(* IEC 61131-3 sources: daoli-st-library/DL_MathData (part 8) *)

(* ---- FC_DL_AngleLerpShort.st ---- *)
(*==============================================================================
 * 名称 : FC_DL_AngleLerpShort —— 两角度最短弧线性插值（跨 0/360 正确）
 * 分类 / 前缀 / 版本 : DL_MathData / FC_DL_ / 1.0.0
 * 溯源 : 开源语义参考（OSCAT/AixOCAT 族，MIT）或 clean-room IEC 实现，未复制源码
 * 平台 : 纯 IEC 61131-3
 * 功能说明 : 沿 fA→fB 最短弧做线性插值：先求 fB-fA 的最短弧差 d∈[-180,180)，
 *            结果 = fA + fT*d，再归一到 [0,360)。fT=0 得 fA 方向，fT=1 得 fB
 *            方向；跨 0/360（如 350°→10°）走 +20° 短弧而非 -340° 长弧。
 *            边界处理：fT 越界 [0,1] 钳位使用（不置故障，属容错钳位）；任一
 *            输入非有限（NaN/±Inf）置 eErr 返回 0.0；|fA|>1.0E12 置 eErr。
 * 错误码 : 16#0001_1B02 = 输入非有限（NaN/±Inf）或角度量超安全量程 ±1.0E12
 *          eErr=0 且 bValid=TRUE 表示返回值可用
 * 状态机 : R6 标注 N/A（纯函数无顺序状态，以本节替代 ELSE 兜底）
 * 红线 : R1/R2/R3 ✓ 零全局/零IO/纯IEC ｜ R4 ✓ 非有限拦截/钳位/量程防护 ｜ R10 ✓ 标准转换 ｜ R11 ✓ 分号收尾 ｜ R15 ✓ 无保留字撞名
 * 修订记录 : 2026-11-23 v1.0.0 首次入库（R76）
 *============================================================================*)
FUNCTION FC_DL_AngleLerpShort : LREAL
VAR_INPUT
    fA : LREAL;    // 插值起点角 [度] / interpolation start angle in degrees
    fB : LREAL;    // 插值终点角 [度] / interpolation end angle in degrees
    fT : LREAL;    // 插值比例 0..1，越界钳位 [无量纲] / interpolation ratio, clamped into [0,1]
END_VAR
VAR_OUTPUT
    eErr   : UDINT;    // 故障码，0=正常，1B02=输入非有限或超量程 / error code
    bError : BOOL;     // TRUE=本件发生故障 / TRUE when fault occurred
    bValid : BOOL;     // TRUE=返回值可用 / TRUE when return value is usable
END_VAR
VAR
    _d : LREAL;        // fA→fB 最短弧差 [度] / shortest-arc diff from A to B
    _n : LREAL;        // 整圈数（TRUNC 截断）[圈] / whole turns via truncation
    _t : LREAL;        // 钳位后的插值比例 [无量纲] / clamped ratio
    _r : LREAL;        // 插值中间结果 [度] / interpolated raw result
END_VAR

FC_DL_AngleLerpShort := 0.0;                 // 返回值预设 0.0 / preset return to zero
eErr   := 16#0000_0000;                      // 故障码清零 / clear error code
bError := FALSE;                             // 故障标志清零 / clear error flag
bValid := TRUE;                              // 预设输出可用 / preset valid flag

IF (fA <> fA) OR ((fA - fA) <> (fA - fA))    // fA 非有限 / fA is NaN or infinite
   OR (fB <> fB) OR ((fB - fB) <> (fB - fB)) // fB 非有限 / fB is NaN or infinite
   OR (fT <> fT) OR ((fT - fT) <> (fT - fT)) // fT 非有限 / fT is NaN or infinite
   OR (ABS(fA) > 1.0E12) OR (ABS(fB) > 1.0E12) THEN    // 角度量超安全量程 / beyond safe range
    eErr   := 16#0001_1B02;                  // 置故障码 / set error code
    bError := TRUE;                          // 置故障标志 / set error flag
    bValid := FALSE;                         // 返回值不可用 / return not usable
    RETURN;                                  // 返回 0.0 / return zero
END_IF

_t := fT;                                    // 取比例 / take ratio
IF _t < 0.0 THEN _t := 0.0; END_IF           // 下界钳位 / clamp lower bound
IF _t > 1.0 THEN _t := 1.0; END_IF           // 上界钳位 / clamp upper bound

_d := fB - fA;                               // 原始差值 / raw difference
_d := _d - 360.0 * TRUNC(_d / 360.0);        // 整圈截断缩圈 / strip whole turns
IF _d >= 180.0 THEN                          // 上越界修正 / fix upper overflow
    _d := _d - 360.0;                        // 减一整圈 / subtract one turn
END_IF
IF _d < -180.0 THEN                          // 下越界修正 / fix lower overflow
    _d := _d + 360.0;                        // 加一整圈 / add one turn
END_IF

_r := fA + _t * _d;                          // 沿最短弧插值 / interpolate along shortest arc
_r := _r - 360.0 * TRUNC(_r / 360.0);        // 归一缩圈 / normalize by stripping turns
IF _r < 0.0 THEN                             // 负角修正 / fix negative angle
    _r := _r + 360.0;                        // 加一整圈 / add one turn
END_IF

FC_DL_AngleLerpShort := _r;                  // 回写 [0,360) 插值结果 / write back result

END_FUNCTION

(* ---- FC_DL_AngleQuadrant.st ---- *)
(*==============================================================================
 * 名称 : FC_DL_AngleQuadrant —— 角度象限判定（0..3）与坐标轴命中标志
 * 分类 / 前缀 / 版本 : DL_MathData / FC_DL_ / 1.0.0
 * 溯源 : 开源语义参考（OSCAT/AixOCAT 族，MIT）或 clean-room IEC 实现，未复制源码
 * 平台 : 纯 IEC 61131-3
 * 功能说明 : 将输入角归一到 [0,360) 后判定象限：0=[0,90) 1=[90,180)
 *            2=[180,270) 3=[270,360)。归一角恰为 0/90/180/270（容差
 *            1.0E-9，浮点禁用 = 直接比较）时 bOnAxis=TRUE，象限取该轴线
 *            后一侧区间编号（0°→0、90°→1、180°→2、270°→3）。
 *            边界处理：输入非有限（NaN/±Inf）或 |角|>1.0E12 置 eErr 返回 0。
 * 错误码 : 16#0001_1B03 = 输入非有限（NaN/±Inf）或角度量超安全量程 ±1.0E12
 *          eErr=0 且 bValid=TRUE 表示象限与轴标志均可用
 * 状态机 : R6 标注 N/A（纯函数无顺序状态，以本节替代 ELSE 兜底）
 * 红线 : R1/R2/R3 ✓ 零全局/零IO/纯IEC ｜ R4 ✓ 非有限拦截/浮点容差比较 ｜ R10 ✓ 标准转换 ｜ R11 ✓ 分号收尾 ｜ R15 ✓ 无保留字撞名
 * 修订记录 : 2026-11-23 v1.0.0 首次入库（R76）
 *============================================================================*)
FUNCTION FC_DL_AngleQuadrant : INT
VAR_INPUT
    fAngle : LREAL;    // 输入角（任意实数，内部归一）[度] / input angle, normalized internally
END_VAR
VAR_OUTPUT
    bOnAxis : BOOL;    // TRUE=归一角命中 0/90/180/270（容差 1.0E-9）/ TRUE when on axis within 1.0E-9
    eErr    : UDINT;   // 故障码，0=正常，1B03=输入非有限或超量程 / error code
    bError  : BOOL;    // TRUE=本件发生故障 / TRUE when fault occurred
    bValid  : BOOL;    // TRUE=象限与轴标志可用 / TRUE when outputs are usable
END_VAR
VAR
    _r : LREAL;        // 归一后的角 [度] / normalized angle
    _n : LREAL;        // 整圈数（TRUNC 截断）[圈] / whole turns via truncation
END_VAR

FC_DL_AngleQuadrant := 0;                    // 象限预设 0 / preset quadrant to zero
bOnAxis := FALSE;                            // 轴标志预设 FALSE / preset on-axis to FALSE
eErr    := 16#0000_0000;                     // 故障码清零 / clear error code
bError  := FALSE;                            // 故障标志清零 / clear error flag
bValid  := TRUE;                             // 预设输出可用 / preset valid flag

IF (fAngle <> fAngle) OR ((fAngle - fAngle) <> (fAngle - fAngle))    // 非有限 / NaN or infinite
   OR (ABS(fAngle) > 1.0E12) THEN            // 超安全量程 / beyond safe range
    eErr   := 16#0001_1B03;                  // 置故障码 / set error code
    bError := TRUE;                          // 置故障标志 / set error flag
    bValid := FALSE;                         // 输出不可用 / outputs not usable
    RETURN;                                  // 返回 0 / return zero
END_IF

_r := fAngle;                                // 取输入角 / take input
_r := _r - 360.0 * TRUNC(_r / 360.0);        // 整圈截断缩圈 / strip whole turns
IF _r < 0.0 THEN                             // 负角修正 / fix negative angle
    _r := _r + 360.0;                        // 加一整圈，得 [0,360) / add one turn
END_IF

IF ABS(_r - 0.0) < 1.0E-9                    // 轴线 0°（含容差）/ on axis 0 deg
   OR ABS(_r - 90.0) < 1.0E-9                // 轴线 90°（含容差）/ on axis 90 deg
   OR ABS(_r - 180.0) < 1.0E-9               // 轴线 180°（含容差）/ on axis 180 deg
   OR ABS(_r - 270.0) < 1.0E-9 THEN          // 轴线 270°（含容差）/ on axis 270 deg
    bOnAxis := TRUE;                         // 置轴线命中标志 / set on-axis flag
END_IF

IF _r >= 270.0 THEN                          // [270,360) 第 4 象限 / quadrant 4
    FC_DL_AngleQuadrant := 3;                // 象限码 3 / quadrant code 3
ELSIF _r >= 180.0 THEN                       // [180,270) 第 3 象限 / quadrant 3
    FC_DL_AngleQuadrant := 2;                // 象限码 2 / quadrant code 2
ELSIF _r >= 90.0 THEN                        // [90,180) 第 2 象限 / quadrant 2
    FC_DL_AngleQuadrant := 1;                // 象限码 1 / quadrant code 1
ELSE                                         // [0,90) 第 1 象限 / quadrant 1
    FC_DL_AngleQuadrant := 0;                // 象限码 0 / quadrant code 0
END_IF

END_FUNCTION

(* ---- FC_DL_AngleReflect.st ---- *)
(*==============================================================================
 * 名称 : FC_DL_AngleReflect —— 关于轴线角 fAxis 的镜像反射（结果 [0,360)）
 * 分类 / 前缀 / 版本 : DL_MathData / FC_DL_ / 1.0.0
 * 溯源 : 开源语义参考（OSCAT/AixOCAT 族，MIT）或 clean-room IEC 实现，未复制源码
 * 平台 : 纯 IEC 61131-3
 * 功能说明 : 求入射角 fAngle 关于镜像轴 fAxis 的反射角：r = 2*fAxis - fAngle
 *            （数值语义恒正确，含跨 0°/360° 情形），归一到 [0,360)。
 *            例：轴 45°、入射 10° → 反射 80°；轴 0°、入射 350° → 反射 10°。
 *            边界处理：任一输入非有限（NaN/±Inf）或 |量|>1.0E12 置 eErr 返回 0.0。
 * 错误码 : 16#0001_1B07 = 输入非有限（NaN/±Inf）或角度量超安全量程 ±1.0E12
 *          eErr=0 且 bValid=TRUE 表示返回值可用
 * 状态机 : R6 标注 N/A（纯函数无顺序状态，以本节替代 ELSE 兜底）
 * 红线 : R1/R2/R3 ✓ 零全局/零IO/纯IEC ｜ R4 ✓ 非有限拦截/量程防护 ｜ R10 ✓ 标准转换 ｜ R11 ✓ 分号收尾 ｜ R15 ✓ 无保留字撞名
 * 修订记录 : 2026-11-23 v1.0.0 首次入库（R76）
 *============================================================================*)
FUNCTION FC_DL_AngleReflect : LREAL
VAR_INPUT
    fAngle : LREAL;    // 入射角 [度] / incident angle in degrees
    fAxis  : LREAL;    // 镜像轴角 [度] / mirror axis angle in degrees
END_VAR
VAR_OUTPUT
    eErr   : UDINT;    // 故障码，0=正常，1B07=输入非有限或超量程 / error code
    bError : BOOL;     // TRUE=本件发生故障 / TRUE when fault occurred
    bValid : BOOL;     // TRUE=返回值可用 / TRUE when return value is usable
END_VAR
VAR
    _r : LREAL;        // 反射角中间值 [度] / reflected raw angle
END_VAR

FC_DL_AngleReflect := 0.0;                   // 返回值预设 0.0 / preset return to zero
eErr   := 16#0000_0000;                      // 故障码清零 / clear error code
bError := FALSE;                             // 故障标志清零 / clear error flag
bValid := TRUE;                              // 预设输出可用 / preset valid flag

IF (fAngle <> fAngle) OR ((fAngle - fAngle) <> (fAngle - fAngle))    // fAngle 非有限 / NaN or infinite
   OR (fAxis <> fAxis) OR ((fAxis - fAxis) <> (fAxis - fAxis))        // fAxis 非有限 / NaN or infinite
   OR (ABS(fAngle) > 1.0E12) OR (ABS(fAxis) > 1.0E12) THEN            // 角度量超安全量程 / beyond safe range
    eErr   := 16#0001_1B07;                  // 置故障码 / set error code
    bError := TRUE;                          // 置故障标志 / set error flag
    bValid := FALSE;                         // 返回值不可用 / return not usable
    RETURN;                                  // 返回 0.0 / return zero
END_IF

_r := 2.0 * fAxis - fAngle;                  // 关于轴镜像反射 / reflect about axis
_r := _r - 360.0 * TRUNC(_r / 360.0);        // 整圈截断缩圈 / strip whole turns
IF _r < 0.0 THEN                             // 负角修正 / fix negative angle
    _r := _r + 360.0;                        // 加一整圈，得 [0,360) / add one turn
END_IF

FC_DL_AngleReflect := _r;                    // 回写 [0,360) 反射角 / write back reflection

END_FUNCTION

(* ---- FC_DL_AngleToCompass.st ---- *)
(*==============================================================================
 * 名称 : FC_DL_AngleToCompass —— 方位角转 16 方位码（0=北，顺时针）与 8 方位码
 * 分类 / 前缀 / 版本 : DL_MathData / FC_DL_ / 1.0.0
 * 溯源 : 开源语义参考（OSCAT/AixOCAT 族，MIT）或 clean-room IEC 实现，未复制源码
 * 平台 : 纯 IEC 61131-3
 * 功能说明 : 将方位角归一到 [0,360) 后按每扇区 22.5° 映射到 16 方位码
 *            0..15（0=北、4=东、8=南、12=西，顺时针），并以 45° 扇区同步
 *            给出 8 方位码 nBand 0..7（0=北、2=东、4=南、6=西），供下游
 *            粗分级直接使用。扇区中心对齐：加半扇区 11.25°/22.5° 后取整。
 *            边界处理：输入非有限（NaN/±Inf）或 |角|>1.0E12 置 eErr 返回 0。
 * 错误码 : 16#0001_1B05 = 输入非有限（NaN/±Inf）或角度量超安全量程 ±1.0E12
 *          eErr=0 且 bValid=TRUE 表示两码均可用
 * 状态机 : R6 标注 N/A（纯函数无顺序状态，以本节替代 ELSE 兜底）
 * 红线 : R1/R2/R3 ✓ 零全局/零IO/纯IEC ｜ R4 ✓ 非有限拦截/量程防护 ｜ R10 ✓ 标准转换 ｜ R11 ✓ 分号收尾 ｜ R15 ✓ 无保留字撞名
 * 修订记录 : 2026-11-23 v1.0.0 首次入库（R76）
 *============================================================================*)
FUNCTION FC_DL_AngleToCompass : INT
VAR_INPUT
    fAngle : LREAL;    // 方位角（0=北，顺时针为正）[度] / bearing angle, clockwise from north
END_VAR
VAR_OUTPUT
    nBand  : INT;      // 8 方位码 0..7（0=北）/ 8-point compass code
    eErr   : UDINT;    // 故障码，0=正常，1B05=输入非有限或超量程 / error code
    bError : BOOL;     // TRUE=本件发生故障 / TRUE when fault occurred
    bValid : BOOL;     // TRUE=两码均可用 / TRUE when both codes are usable
END_VAR
VAR
    _r    : LREAL;     // 归一后的方位角 [度] / normalized bearing
    _n16  : LREAL;     // 16 扇区整数值 / 16-sector integer value
    _n8   : LREAL;     // 8 扇区整数值 / 8-sector integer value
END_VAR

FC_DL_AngleToCompass := 0;                   // 16 码预设 0（北）/ preset 16-code to north
nBand := 0;                                  // 8 码预设 0（北）/ preset 8-code to north
eErr  := 16#0000_0000;                       // 故障码清零 / clear error code
bError:= FALSE;                              // 故障标志清零 / clear error flag
bValid:= TRUE;                               // 预设输出可用 / preset valid flag

IF (fAngle <> fAngle) OR ((fAngle - fAngle) <> (fAngle - fAngle))    // 非有限 / NaN or infinite
   OR (ABS(fAngle) > 1.0E12) THEN            // 超安全量程 / beyond safe range
    eErr   := 16#0001_1B05;                  // 置故障码 / set error code
    bError := TRUE;                          // 置故障标志 / set error flag
    bValid := FALSE;                         // 输出不可用 / outputs not usable
    RETURN;                                  // 返回 0 / return north codes
END_IF

_r := fAngle;                                // 取输入角 / take input
_r := _r - 360.0 * TRUNC(_r / 360.0);        // 整圈截断缩圈 / strip whole turns
IF _r < 0.0 THEN                             // 负角修正 / fix negative angle
    _r := _r + 360.0;                        // 加一整圈，得 [0,360) / add one turn
END_IF

_n16 := TRUNC((_r + 11.25) / 22.5);          // 16 扇区中心对齐取整 / 16-sector center-aligned
_n8  := TRUNC((_r + 22.5) / 45.0);           // 8 扇区中心对齐取整 / 8-sector center-aligned

FC_DL_AngleToCompass := DINT_TO_INT(LREAL_TO_DINT(_n16) MOD 16);    // 折回 0..15 / fold into 0..15
nBand := DINT_TO_INT(LREAL_TO_DINT(_n8) MOD 8);           // 折回 0..7 / fold into 0..7

END_FUNCTION

(* ---- FC_DL_AngleTolInside.st ---- *)
(*==============================================================================
 * 名称 : FC_DL_AngleTolInside —— 角度容差窗判定（fCenter ± fTol，跨 0° 正确）
 * 分类 / 前缀 / 版本 : DL_MathData / FC_DL_ / 1.0.0
 * 溯源 : 开源语义参考（OSCAT/AixOCAT 族，MIT）或 clean-room IEC 实现，未复制源码
 * 平台 : 纯 IEC 61131-3
 * 功能说明 : 判定 fAngle 是否落在 fCenter ± fTol 的圆周窗内：取 fAngle-fCenter
 *            的最短弧差 d∈[-180,180)（天然跨 0°/360° 正确），当 |d| <= fTol
 *            判在内。窗宽 >180° 时窗覆盖超过半圆，仍按最短弧口径判定。
 *            边界处理：fTol<0 判参数非法（置 eErr 返回 FALSE）；任一角度输入
 *            非有限（NaN/±Inf）或 |角|>1.0E12 置 eErr 返回 FALSE。
 * 错误码 : 16#0001_1B06 = fTol 为负（容差非法），或角度输入非有限 / 超安全量程 ±1.0E12
 *          eErr=0 且 bValid=TRUE 表示判定结论可用
 * 状态机 : R6 标注 N/A（纯函数无顺序状态，以本节替代 ELSE 兜底）
 * 红线 : R1/R2/R3 ✓ 零全局/零IO/纯IEC ｜ R4 ✓ 非有限拦截/浮点容差比较 ｜ R10 ✓ 标准转换 ｜ R11 ✓ 分号收尾 ｜ R15 ✓ 无保留字撞名
 * 修订记录 : 2026-11-23 v1.0.0 首次入库（R76）
 *============================================================================*)
FUNCTION FC_DL_AngleTolInside : BOOL
VAR_INPUT
    fAngle  : LREAL;   // 被判定角 [度] / angle under test in degrees
    fCenter : LREAL;   // 窗中心角 [度] / window center angle in degrees
    fTol    : LREAL;   // 容差半窗宽，须 >=0 [度] / tolerance half-width, must be >= 0
END_VAR
VAR_OUTPUT
    eErr   : UDINT;    // 故障码，0=正常，1B06=参数非法或非有限 / error code
    bError : BOOL;     // TRUE=本件发生故障 / TRUE when fault occurred
    bValid : BOOL;     // TRUE=判定结论可用 / TRUE when verdict is usable
END_VAR
VAR
    _d : LREAL;        // 最短弧差 [度] / shortest-arc diff
END_VAR

FC_DL_AngleTolInside := FALSE;               // 判定预设 FALSE / preset verdict to FALSE
eErr   := 16#0000_0000;                      // 故障码清零 / clear error code
bError := FALSE;                             // 故障标志清零 / clear error flag
bValid := TRUE;                              // 预设输出可用 / preset valid flag

IF fTol < 0.0 THEN                           // 容差为负：参数非法 / negative tolerance invalid
    eErr   := 16#0001_1B06;                  // 置参数非法码 / set invalid-parameter code
    bError := TRUE;                          // 置故障标志 / set error flag
    bValid := FALSE;                         // 结论不可用 / verdict not usable
    RETURN;                                  // 返回 FALSE / return FALSE
END_IF

IF (fAngle <> fAngle) OR ((fAngle - fAngle) <> (fAngle - fAngle))     // fAngle 非有限 / NaN or infinite
   OR (fCenter <> fCenter) OR ((fCenter - fCenter) <> (fCenter - fCenter))   // fCenter 非有限 / NaN or infinite
   OR (fTol <> fTol) OR ((fTol - fTol) <> (fTol - fTol))               // fTol 非有限 / NaN or infinite
   OR (ABS(fAngle) > 1.0E12) OR (ABS(fCenter) > 1.0E12) THEN           // 角度量超安全量程 / beyond safe range
    eErr   := 16#0001_1B06;                  // 置故障码 / set error code
    bError := TRUE;                          // 置故障标志 / set error flag
    bValid := FALSE;                         // 结论不可用 / verdict not usable
    RETURN;                                  // 返回 FALSE / return FALSE
END_IF

_d := fAngle - fCenter;                      // 原始差值 / raw difference
_d := _d - 360.0 * TRUNC(_d / 360.0);        // 整圈截断缩圈 / strip whole turns
IF _d >= 180.0 THEN                          // 上越界修正 / fix upper overflow
    _d := _d - 360.0;                        // 减一整圈 / subtract one turn
END_IF
IF _d < -180.0 THEN                          // 下越界修正 / fix lower overflow
    _d := _d + 360.0;                        // 加一整圈 / add one turn
END_IF

IF ABS(_d) <= fTol THEN                      // 最短弧差落在容差窗内 / diff inside tolerance window
    FC_DL_AngleTolInside := TRUE;            // 判在内 / verdict inside
END_IF

END_FUNCTION

(* ---- FC_DL_AngleUnwrapStep.st ---- *)
(*==============================================================================
 * 名称 : FC_DL_AngleUnwrapStep —— 增量解卷绕（跨多圈连续跟踪，步进 [-180,180)）
 * 分类 / 前缀 / 版本 : DL_MathData / FC_DL_ / 1.0.0
 * 溯源 : 开源语义参考（OSCAT/AixOCAT 族，MIT）或 clean-room IEC 实现，未复制源码
 * 平台 : 纯 IEC 61131-3
 * 功能说明 : 编码器增量解卷绕：取 fRaw-fPrev 的最短弧差作为本拍步进
 *            fStep∈[-180,180)，返回 fAccum + fStep 的累计角（不卷绕、跨多圈
 *            连续跟踪）。调用方须把返回值与 fStep 存为下一拍的 fAccum/fPrev。
 *            边界处理：任一输入非有限（NaN/±Inf）或 |量|>1.0E12 置 eErr
 *            返回 fAccum 原值（冻结本拍步进，不引入伪增量）。
 * 错误码 : 16#0001_1B08 = 输入非有限（NaN/±Inf）或角度量超安全量程 ±1.0E12
 *          eErr=0 且 bValid=TRUE 表示步进与累计角均可用
 * 状态机 : R6 标注 N/A（纯函数无顺序状态，跨拍状态由调用方持有，以本节替代 ELSE 兜底）
 * 红线 : R1/R2/R3 ✓ 零全局/零IO/纯IEC ｜ R4 ✓ 非有限拦截/量程防护 ｜ R10 ✓ 标准转换 ｜ R11 ✓ 分号收尾 ｜ R15 ✓ 无保留字撞名
 * 修订记录 : 2026-11-23 v1.0.0 首次入库（R76）
 *============================================================================*)
FUNCTION FC_DL_AngleUnwrapStep : LREAL
VAR_INPUT
    fRaw   : LREAL;    // 本拍原始角 [度] / raw angle of this cycle
    fPrev  : LREAL;    // 上一拍原始角（调用方持有）[度] / previous raw angle, caller-held
    fAccum : LREAL;    // 累计角（调用方持有）[度] / accumulated angle, caller-held
END_VAR
VAR_OUTPUT
    fStep  : LREAL;    // 本拍步进 [-180,180) [度] / step of this cycle within [-180,180)
    eErr   : UDINT;    // 故障码，0=正常，1B08=输入非有限或超量程 / error code
    bError : BOOL;     // TRUE=本件发生故障 / TRUE when fault occurred
    bValid : BOOL;     // TRUE=步进与累计角可用 / TRUE when step and result are usable
END_VAR
VAR
    _d : LREAL;        // 本拍原始差值 [度] / raw delta of this cycle
END_VAR

fStep := 0.0;                                // 步进预设 0.0 / preset step to zero
eErr   := 16#0000_0000;                      // 故障码清零 / clear error code
bError := FALSE;                             // 故障标志清零 / clear error flag
bValid := TRUE;                              // 预设输出可用 / preset valid flag
FC_DL_AngleUnwrapStep := fAccum;             // 返回值预设为累计角原值 / preset return to accum

IF (fRaw <> fRaw) OR ((fRaw - fRaw) <> (fRaw - fRaw))      // fRaw 非有限 / NaN or infinite
   OR (fPrev <> fPrev) OR ((fPrev - fPrev) <> (fPrev - fPrev))   // fPrev 非有限 / NaN or infinite
   OR (fAccum <> fAccum) OR ((fAccum - fAccum) <> (fAccum - fAccum))  // fAccum 非有限 / NaN or infinite
   OR (ABS(fRaw) > 1.0E12) OR (ABS(fPrev) > 1.0E12) THEN     // 角度量超安全量程 / beyond safe range
    eErr   := 16#0001_1B08;                  // 置故障码 / set error code
    bError := TRUE;                          // 置故障标志 / set error flag
    bValid := FALSE;                         // 输出不可用 / outputs not usable
    RETURN;                                  // 冻结本拍，返回 fAccum 原值 / freeze, return accum unchanged
END_IF

_d := fRaw - fPrev;                          // 本拍原始差值 / raw delta
_d := _d - 360.0 * TRUNC(_d / 360.0);        // 整圈截断缩圈 / strip whole turns
IF _d >= 180.0 THEN                          // 上越界修正（取短弧步进）/ fix upper overflow
    _d := _d - 360.0;                        // 减一整圈 / subtract one turn
END_IF
IF _d < -180.0 THEN                          // 下越界修正 / fix lower overflow
    _d := _d + 360.0;                        // 加一整圈 / add one turn
END_IF

fStep := _d;                                 // 回写本拍步进 / write back step
FC_DL_AngleUnwrapStep := fAccum + _d;        // 累计角连续跟踪（不卷绕）/ accumulate unwrapped

END_FUNCTION

(* ---- FC_DL_AnodizeFilmThicknessCalc.st ---- *)
(*
  Component : FC_DL_AnodizeFilmThicknessCalc
  Category  : DL_MathData
  Type      : FC
  Complexity: C1
  VERSION   : v1.0.0
  功能      : 阳极氧化膜厚-电量换算：按法拉第定律由电量密度与膜密度算膜厚 μm，并按电流密度反算达目标膜厚所需时间。
  开源溯源  : 道莅原创 clean-room 自研（无外部代码引用）｜License: MIT
  边界条件  : ① 膜密度、摩尔质量、转移电子数须 > 1e-9，效率须在 (0,100] % 内，否则返回哨兵 -1；
              ② 反算时间需电流密度 > 1e-9，电流密度为 0 时时间回 0（不下发 inf）；
              ③ 量纲链：g/dm² ÷ g/cm³ = cm³/dm²，除 dm² 面积 100 cm² 得 cm 厚，再乘 1e4 得 μm。
*)
FUNCTION FC_DL_AnodizeFilmThicknessCalc : REAL
VAR_INPUT
    fChgDensAsDm2 : REAL;   (* 电量密度 [A·s/dm²] Charge density *)
    fMolarMassGmol: REAL;   (* 氧化物摩尔质量 [g/mol] Oxide molar mass *)
    fDensityGcm3  : REAL;   (* 膜层密度 [g/cm³] Film density *)
    nElectrons    : INT;    (* 反应转移电子数 [个] Transferred electrons *)
    fEffPct       : REAL;   (* 电流效率 [%] Current efficiency *)
    fCurrDensADm2 : REAL;   (* 电流密度 [A/dm²] Current density *)
    fThickTargetUm: REAL;   (* 目标膜厚 [μm] Target film thickness *)
END_VAR
VAR_OUTPUT
    fFilmUm        : REAL;  (* 膜厚 [μm] Film thickness *)
    fMassGdm2      : REAL;  (* 单位面积氧化膜质量 [g/dm²] Film mass per area *)
    fTimeForTargetS: REAL;  (* 达目标膜厚所需时间 [s] Time to reach target thickness *)
    xValid         : BOOL;  (* 计算有效性标志 [-] Calculation valid flag *)
END_VAR
VAR CONSTANT
    DL_EPS      : REAL := 1.0E-9;   (* 除零判定容差 [无量纲] Divide-by-zero tolerance *)
    DL_FARADAY  : REAL := 96485.332;(* 法拉第常数 [C/mol] Faraday constant *)
    DL_CM_PER_DM: REAL := 100.0;    (* dm² 对应 cm² 数 [cm²/dm²] cm2 per dm2 *)
    DL_PCT_BASE : REAL := 100.0;    (* 百分比基准 [%] Percent base *)
    DL_UM_PER_CM: REAL := 10000.0;  (* 厘米转微米系数 [μm/cm] Micrometres per centimetre *)
    DL_ZERO     : REAL := 0.0;      (* 零常量 [无量纲] Zero constant *)
END_VAR
VAR
    fEffUnit : REAL;   (* 效率折算系数 [-] Efficiency as fraction *)
    fMoles   : REAL;   (* 单位面积反应摩尔数 [mol/dm²] Moles per area *)
END_VAR
(* 出口预置：四出口统一预置 *)
fFilmUm := 0.0; fMassGdm2 := 0.0; fTimeForTargetS := 0.0; xValid := FALSE;
(* 非有限拦截：自反判 NaN，自身差值判 Inf *)
IF (fChgDensAsDm2 <> fChgDensAsDm2) OR ((fChgDensAsDm2 - fChgDensAsDm2) <> 0.0)
   OR (fMolarMassGmol <> fMolarMassGmol) OR ((fMolarMassGmol - fMolarMassGmol) <> 0.0)
   OR (fDensityGcm3 <> fDensityGcm3) OR ((fDensityGcm3 - fDensityGcm3) <> 0.0)
   OR (fEffPct <> fEffPct) OR ((fEffPct - fEffPct) <> 0.0)
   OR (fCurrDensADm2 <> fCurrDensADm2) OR ((fCurrDensADm2 - fCurrDensADm2) <> 0.0) THEN
    FC_DL_AnodizeFilmThicknessCalc := -1.0;  (* 哨兵 -1：输入非有限 / Sentinel -1 non-finite *)
    RETURN;
END_IF
(* 组态域闸：膜密度、摩尔质量、转移电子数、效率、电量密度非负 *)
IF (fDensityGcm3 <= DL_EPS) OR (fMolarMassGmol <= DL_EPS) OR (nElectrons < 1)
   OR (fEffPct <= DL_ZERO) OR (fEffPct > DL_PCT_BASE) OR (fChgDensAsDm2 < DL_ZERO) THEN
    FC_DL_AnodizeFilmThicknessCalc := -1.0;  (* 哨兵 -1：组态非法 / Sentinel -1 bad config *)
    RETURN;
END_IF
fEffUnit := fEffPct / DL_PCT_BASE;             (* 效率折算 [-] / Efficiency as fraction *)
(* 单位面积摩尔数：n = q / (z·F)，电量密度为 C/dm² *)
fMoles := fChgDensAsDm2 / (INT_TO_REAL(nElectrons) * DL_FARADAY);
(* 单位面积质量：m = n·M [g/dm²]，乘效率得实际成膜量 *)
fMassGdm2 := fMoles * fMolarMassGmol * fEffUnit;
(* 厚度换算：g/dm² ÷ g/cm³ = cm³/dm²，除 100 cm² 得 cm，再乘 1e4 得 μm *)
fFilmUm := (fMassGdm2 / fDensityGcm3) / DL_CM_PER_DM * DL_UM_PER_CM;
(* 反算时间：t = 目标膜厚 / (电流密度 × 单位电量膜厚系数)，电流密度为 0 时回 0 *)
IF (fCurrDensADm2 > DL_EPS) AND (fThickTargetUm > DL_ZERO) THEN
    fTimeForTargetS := fThickTargetUm * INT_TO_REAL(nElectrons) * DL_FARADAY * fDensityGcm3
                       / (fCurrDensADm2 * fMolarMassGmol * fEffUnit * DL_CM_PER_DM);
END_IF
xValid := TRUE;                                (* 链路有效 / Chain valid *)
FC_DL_AnodizeFilmThicknessCalc := fFilmUm;     (* 返回膜厚 [μm] / Return film thickness *)
END_FUNCTION

(* ---- FC_DL_ArrayCumSumLreal.st ---- *)
(*
    FC_DL_ArrayCumSumLreal —— LREAL 数组前缀累计序列 + 总和出口（统计线）
    ------------------------------------------------------------------
    组件名称  : FC_DL_ArrayCumSumLreal
    分类      : DL_MathData / Statistics
    前缀      : FC_DL_
    版本      : 1.0.0
    溯源      : 借鉴组织 —— T2-1 LGF · Math（统计线，矩阵行 157）：仅借鉴
                「前缀累计 / 累计序列输出」公开功能定义；clean-room 声明 ——
                零代码行复制，判据链 / 码位 / 钳位与拒绝口径 100% 自有；
                累加内核为 IEC 61131-3 标准算术的道莅防御性实现。
    平台      : 纯 IEC 61131-3（WHILE + LREAL 算术），无内建函数依赖，
                CODESYS 3.5 / TwinCAT 3 / InoProShop / Machine Expert 通用
    作者      : 道莅代码库 · PLC编程专家（R72 构建轮 · 批 1 · 序号 3）
    ------------------------------------------------------------------
    功能说明  : 对有效样本数 nCount 个 LREAL 输入计算前缀累计序列
                afOut[i] = Σ afIn[1..i]（i = 1..nCount），并给总和出口
                fTotal = afOut[nCount]。真实工况：能耗 / 产量累计曲线、
                按片批次余量推演、OEE 累计谱。量纲随输入（m³ / kWh / 件 等），
                本件不解释量纲。
                判据链顺序：
                ① nCount 域闸：0 → 信息级空出口（fTotal = 0，afOut 不触碰，
                   bValid = TRUE）；> 数组上界 → 钳位照算 + 信息级；
                ② 逐元素非有限闸（两遍扫描第一遍，R151 闸全枚举）：**遇非有限
                   样本整体拒绝**（保守口径：部分累计会污染下游余量判断，
                   出故障级码，afOut 零写入）；
                ③ 循环累加（WHILE 带 DL_CUM_GUARD 防死锁计数器，两遍各自独立
                   计数）+ 写前下标双检；
                ④ 溢出面：累计 > 1E30 → 置 bTruncated 中断累加（保留至上一
                   有效前缀），信息级声明口径；非有限中间量同判（差值自反 +
                   自反双判，R79）。
                浮点判等禁用 =（红线 5）：本件无浮点相等比较。
    错误码    : 16#0002_3902 nCount = 0，空出口（fTotal = 0，bValid = TRUE）
                            —— 信息级，不置 bError（R45）
                16#0002_3903 nCount > 数组上界，已钳位照算 —— 信息级，值可用
                16#0002_3904 样本非有限或循环守卫越限（整体拒绝，afOut 零写入，
                            返回 FALSE）—— 故障级
                16#0002_3905 累计超 1E30 上界，已置 bTruncated 中断累加（保留
                            至上一有效前缀，bValid = TRUE）—— 信息级
                加码反证句（R90）：3902/3903/3905 均有独立输出观测面
                （3902 由 nCount=0 请求 + 空出口唯一对应；3903 由钳位行为 +
                部分结果唯一对应；3905 由 bTruncated 专位唯一对应），互不可
                由现有输出组合还原，故各立一码。
    码位总账  : 16#0002_3902 用 ｜ 16#0002_3903 用 ｜ 16#0002_3904 用 ｜
                16#0002_3905 用
    状态机    : N/A —— 纯函数无状态，无 CASE 可写，非法状态不可能出现
    边界与披露: 一 无定时器 / 无沿检测实例，周期安全规则 N/A；WHILE 双循环
                   各配 DL_CUM_GUARD 守卫（160 > 上界 128，正常不触发），
                   守卫越限并入 3904 故障级（结构性不可达防御收口）；
                二 零全局变量、零 VAR_EXTERNAL、零物理地址；
                三 域闸逐项点名（R272）：afIn[1..nEff] 全部元素纳入非有限闸；
                   nCount 域闸覆盖 0 / 上界两端点（各推一条向量）；
                四 数组写前下标双检（红线 2）：(nI >= 1) AND (nI <= DL_CUM_NMAX)
                   显式兜底；下标 > nCount 的 afOut 元素不被本件触碰；
                五 除法面：无（零除法，零除零面）；
                六 与 FC_DL_ArraySumLreal（DL_MathData）分工互引：后者只出
                   总和（可零拷贝、非有限剔除口径），本件输出**完整前缀序列**
                   （须写入调用方数组、整体拒绝口径），非变体，分工写死。
    验收向量  : V1 afIn = [1,2,3]，nCount = 3 → afOut = [1,3,6]，fTotal = 6；
                V2 nCount = 0 → 空出口 3902，fTotal = 0，afOut 不触碰；
                V3 nCount = 200（> 128）→ 钳位照算 3903；
                V4 afIn[2] = NaN → 3904 故障级，afOut 零写入；
                V5 累计越 1E30 → bTruncated = TRUE + 3905。
                算法已证（脚本）：未跑 ｜ 编译器已证（三平台）：未跑
    修订记录  : 2026-11-23 v1.0.0 首次入库（R72 构建轮 · 批 1 · 序号 3）
*)
FUNCTION FC_DL_ArrayCumSumLreal : BOOL
VAR_INPUT
    nCount    : UDINT;                     (* 有效样本数，[个]，0 = 空出口，超上界钳位照算 / the valid sample count *)
END_VAR
VAR_IN_OUT
    afIn      : ARRAY[1..DL_CUM_NMAX] OF LREAL;  (* 输入样本数组，[量纲随输入]，下标 1 起 / the input samples, unit follows the caller *)
    afOut     : ARRAY[1..DL_CUM_NMAX] OF LREAL;  (* 前缀累计序列出口，[量纲随输入]，afOut[i] = Σ afIn[1..i] / the prefix cumulative output *)
END_VAR
VAR_OUTPUT
    fTotal     : LREAL;                    (* 总和出口 = afOut[nCount]（截断时为最后有效前缀），[量纲随输入] / the total outlet *)
    bTruncated : BOOL;                     (* 累计越 1E30 上界截断标志 / the truncation flag *)
    bValid     : BOOL;                     (* 输出可用标志，故障级为 FALSE / the outputs usable flag *)
    bError     : BOOL;                     (* 故障标志，仅故障级码置位（R45 配对）/ the fault flag *)
    nInfoCode  : UDINT;                    (* 信息 / 错误码，0 = 正常 / the info or error id *)
END_VAR
VAR CONSTANT
    DL_CUM_NMAX  : INT  := 128;            (* 数组上界（两数组维度必须与本常量一致）[个] / the array upper bound, both arrays must match *)
    DL_CUM_NMAXU : UDINT := 128;           (* 数组上界的 UDINT 影子（nCount 域闸同口径比较用）[个] / the UDINT shadow of the bound *)
    DL_CUM_CAP   : LREAL := 1.0E30;        (* 累计幅值上界（截断口径）[量纲随输入] / the cumulative magnitude cap *)
    DL_CUM_GUARD : INT  := 160;            (* 循环守卫上限（> 上界 128，正常不触发）[次] / the loop guard limit *)
    DL_CUM_ZERO  : LREAL := 0.0;           (* 零哨兵 [量纲随输入] / the zero sentinel *)
    DL_CUM_ONE   : INT  := 1;              (* 游标步进与下界常量 [个] / the cursor step and lower bound *)
END_VAR
VAR
    nEff    : INT;                         (* 钳位后的有效样本数 [个] / the effective clamped count *)
    nI      : INT;                         (* 数组游标 [个] / the array cursor *)
    nGuard  : INT;                         (* 循环守卫计数器 [次] / the loop guard counter *)
    fRun    : LREAL;                       (* 累加器 [量纲随输入] / the running accumulator *)
    bFinOk  : BOOL;                        (* 第一遍有限性扫描结论 / the pass one finiteness verdict *)
    bStop   : BOOL;                        (* 第二遍截断中止标志 / the pass two truncation stop flag *)
    bSmpFin : BOOL;                        (* 当前样本有限性中间结论 / the per sample finiteness temporary *)
END_VAR

// 段 1｜返回值与状态预置（统一出口预置，R256）/ segment 1, preset the return and the status
FC_DL_ArrayCumSumLreal := FALSE;         // 故障缺省返回不可用 / the fault default is unusable
fTotal     := DL_CUM_ZERO;               // 总和出口预置零 / preset the total to zero
bTruncated := FALSE;                     // 截断标志预清零 / preset the truncation flag false
bValid     := FALSE;                     // 可用标志预清零 / preset the usable flag false
bError     := FALSE;                     // 故障标志预清零 / preset the fault flag false
nInfoCode  := 0;                         // 码位预置无错 / preset the code to zero
nEff    := 0;                            // 有效数预置零 / preset the effective count zero
nI      := 0;                            // 游标预置零 / preset the cursor zero
nGuard  := 0;                            // 守卫预置零 / preset the guard zero
fRun    := DL_CUM_ZERO;                  // 累加器清零 / clear the accumulator
bFinOk  := TRUE;                         // 有限性结论预置通过 / preset the finiteness verdict pass
bStop   := FALSE;                        // 截断标志预清零 / preset the stop flag false
bSmpFin := TRUE;                         // 样本有限性预置通过 / preset the per sample verdict pass

// 段 2｜nCount 域闸（0 = 空出口，超界 = 钳位照算，两端点向量）/ segment 2, the count domain gate
IF nCount = 0 THEN                       // 空请求：信息级空出口（afOut 不触碰）/ an empty request, the empty outlet
    nInfoCode := 16#0002_3902;           // 信息级：空出口 / info level: the empty outlet
    bError := FALSE;                     // 信息级不置故障（R45）/ info level never raises a fault
    bValid := TRUE;                      // 空出口按契约可用 / the empty outlet usable by contract
    FC_DL_ArrayCumSumLreal := TRUE;      // 照算完成（空）/ the pass complete, empty
    RETURN;                              // 结构早退 / structural exit
END_IF
IF nCount > DL_CUM_NMAXU THEN            // 请求超数组上界：钳位照算 / the request over the bound, clamped
    nInfoCode := 16#0002_3903;           // 信息级：已钳位照算 / info level: clamped
    nEff := DL_CUM_NMAX;                 // 钳到上界 / clamp to the bound
ELSE                                     // 域内请求 / the in domain request
    nEff := UDINT_TO_DINT(nCount);       // 降位转换（已证 <= 128，无回绕面）/ the narrowing conversion proven safe
END_IF

// 段 3｜第一遍：逐元素非有限扫描（整体拒绝口径，闸前零写入）/ segment 3, the pass one finiteness scan
nI     := DL_CUM_ONE;                    // 游标从下标 1 起 / the cursor from index one
nGuard := 0;                            // 守卫清零 / clear the guard
WHILE (nI <= nEff) AND (nGuard < DL_CUM_GUARD) DO // 守卫内扫描 / the scan inside the guard
    IF (nI >= DL_CUM_ONE) AND (nI <= DL_CUM_NMAX) THEN // 写前读前下标双检（红线 2）/ the index double check
        bSmpFin := NOT ((afIn[nI] <> afIn[nI]) OR ((afIn[nI] - afIn[nI]) <> 0.0)); // 自反 + 差值自反双判（R79）/ the reflexive pair test
        IF NOT bSmpFin THEN              // 非有限样本命中 / a non finite sample hit
            bFinOk := FALSE;             // 整体拒绝结论 / the overall reject verdict
            nI := nEff + DL_CUM_ONE;     // 跳出扫描（守卫内合法退出）/ break the scan legally
        END_IF
    END_IF
    nI := nI + DL_CUM_ONE;               // 游标推进 / advance the cursor
    nGuard := nGuard + DL_CUM_ONE;       // 守卫推进 / advance the guard
END_WHILE
IF (NOT bFinOk) OR (nGuard >= DL_CUM_GUARD) THEN // 非有限命中或守卫越限 / a hit or a guard overflow
    nInfoCode := 16#0002_3904;           // 故障级：样本序列不可信整体拒绝（守卫越限为结构性不可达防御收口）/ fault level: the samples untrusted
    bError := TRUE;                      // R45 配对置故障标志 / paired with the fault flag
    bValid := FALSE;                     // 输出不可用 / the outputs unusable
    FC_DL_ArrayCumSumLreal := FALSE;     // 拒绝返回 / the reject return
    RETURN;                              // 结构早退（afOut 保持零写入）/ exit with afOut untouched
END_IF

// 段 4｜第二遍：前缀累计与写出口（截断口径：累计 > 1E30 中断累加）/ segment 4, the pass two prefix accumulation
nI     := DL_CUM_ONE;                    // 游标复位 / reset the cursor
nGuard := 0;                             // 守卫复位 / reset the guard
WHILE (nI <= nEff) AND (nGuard < DL_CUM_GUARD) AND (NOT bStop) DO // 守卫与截断双出口 / the loop with both exits
    IF (nI >= DL_CUM_ONE) AND (nI <= DL_CUM_NMAX) THEN // 写前下标双检（红线 2）/ the index double check
        fRun := fRun + afIn[nI];         // 前缀累加（样本已过第一遍闸）/ the prefix accumulation
        IF (fRun <> fRun) OR ((fRun - fRun) <> 0.0) OR (fRun > DL_CUM_CAP) THEN // 溢出面：非有限中间量或越上界 / the overflow surface
            bTruncated := TRUE;          // 置截断标志 / raise the truncation flag
            nInfoCode := 16#0002_3905;   // 信息级：已截断（优先级高于钳位码 3903，声明口径）/ info level: truncated, overriding the clamp code
            bStop := TRUE;               // 中断累加（保留至上一有效前缀）/ stop the accumulation
        ELSE                             // 前缀有效 / the prefix valid
            afOut[nI] := fRun;           // 写前缀出口 / write the prefix outlet
        END_IF
    END_IF
    nI := nI + DL_CUM_ONE;               // 游标推进 / advance the cursor
    nGuard := nGuard + DL_CUM_ONE;       // 守卫推进 / advance the guard
END_WHILE

// 段 5｜正常出口 / segment 5, the normal outlet
fTotal := fRun;                          // 总和出口 = 最后有效前缀 / the total outlet, the last valid prefix
bError := FALSE;                         // 信息级不置故障（双保险）/ info level never raises a fault, second line
bValid := TRUE;                          // 输出可用 / the outputs usable
FC_DL_ArrayCumSumLreal := TRUE;          // 照算完成 / the pass complete
END_FUNCTION

(* ---- FC_DL_ArrayDiffSummary.st ---- *)
(*==============================================================================
 * 组件名称 (Component)  : FC_DL_ArrayDiffSummary
 * 所属子库 (Sublibrary) : DL_MathData
 * 归属目录 (Directory)  : C:\Library\DL_MathData
 * 当前版本 (Version)    : 1.0.1
 * 组件分类 (Category)   : 函数（FUNCTION）· 纯函数 · 双数组逐项容差比对
 * 兼容性   (Platform)   : CODESYS 3.5 / TwinCAT 3 / 汇川 InoProShop / 施耐德
 *                         Machine Expert；仅用 Standard.library 的 ABS，无实例依赖
 * 功能一句话 (Summary)  : 两组实数数组按统一绝对容差逐项比对，输出超差项数、首个
 *                         超差下标、最大绝对偏差及其下标与一致性结论。
 * 功能描述 (Function)   : 配方回读、双通道冗余比对、视觉参数下发校验三类场景，
 *                         现场只判「有差异」却定位不到第几项、差多少；用等号判等
 *                         又会因浮点误差把合格品报成不合格。本件一次扫描给出
 *                         计数、首个位置、最大偏差位置三个定位量，维修工直接翻表。
 * 与既有件边界 (Boundary): FC_DL_SearchMinMax 在单数组内找极值；FC_DL_ArraySearchFirst
 *                         在单数组内按判据找首个命中；本件是双数组逐项配对比较，
 *                         输出统计族，三者职责互斥，不存在覆盖关系。
 * 设计要点 (Key notes)  : ① 容差先取绝对值再钳到最小容差，杜绝「容差为零把纯浮点
 *                           噪声全判超差」的静默失效；
 *                         ② 非数与非有限值前置拦截：该项直接计为超差且不参与最大
 *                           偏差竞争，防止无穷大污染统计结果；
 *                         ③ 最大偏差并列时取先出现者，保证结果可复现；
 *                         ④ 单趟循环完成全部判定，无嵌套循环、无排序、无中间数组；
 *                         ⑤ 纯函数：无内部状态，同入参同结果，可重入。
 * 开源溯源 (Origin)     : 来源标签 lgf-comparator。LGF 为免费闭源发布的公开函数库
 *                         手册，本件仅借鉴其比较器组把「数组批量比较」与「容差窗口」
 *                         分成两个子域的分类骨架；许可证按其发布方条款仅作分类参考，
 *                         本件零代码行、零注释引用，属 clean-room 独立实现。统计口径
 *                         （最大偏差及其下标）为本库自有，LGF 批量比较不输出该量。
 * 码位说明 (Codes)      : 本件独占信息级码段 16#0001_0134 到 16#0001_0135，纯函数
 *                         无锁存面故不占故障级码；与 MathData 既有 0101 到 0124
 *                         及同轮 0125 到 013C 求差为空。
 *                         0134 项数越界已钳位 ｜ 0135 容差非法已回退。
 * 依赖说明 (Depends)    : 无 DL_ 内部依赖；仅 Standard.library 的 ABS。
 * 契约前置条件 (Contract): 函数内无法探测数组实际长度，「nCount 不得大于调用方实际
 *                         数组长度」由调用方负责，组态时须与装载行数绑定。
 * 红线自检 (Redline)    : 零全局变量表依赖 ｜ 零外部变量声明 ｜ 零物理地址
 *                         纯 IEC 61131-3 ｜ 浮点无等号判等，全部走容差 ｜ 无除法
 *                         数组下标先钳位后使用 ｜ 循环带守卫 ｜ 全变量双语同行注释
 * 修订历史 (Revision)   : 2026-11-15  v1.0.0  首版入库（Round 12 · 双数组比对族）
 *                         2026-11-15  v1.0.1  终审定点修复 A-D04：两项有限值相减仍可能
 *                         溢出为无穷（同号异号近满量程），原实现会让该偏差直接参与最大
 *                         偏差竞争并把 fMaxDev 污染成无穷；补「偏差本身超有限上限即按非
 *                         有限处置、不参与竞争」判据，兑现设计要点②的承诺
 *============================================================================*)

(*==============================================================================
 * 比对示意 (Comparison picture)：
 *   期望 10.0 / 20.0 / 30.0，实际 10.0 / 20.005 / 30.2，容差 0.01
 *   第 2 项偏差 0.005 在容差内，合格，但仍是目前最大偏差
 *   第 3 项偏差 0.2 超出容差，超差计数加一，并顶替最大偏差
 *   最终：超差一项、首个超差下标 3、最大偏差 0.2 落在下标 3、不相等
 *   若把实际第 2 项置为非数，该项计为超差且不参与最大偏差竞争
 *============================================================================*)

FUNCTION FC_DL_ArrayDiffSummary : BOOL
VAR_IN_OUT
    afExpected : ARRAY[1..64] OF REAL;   // 期望值数组，基准侧，只读不写 [工程单位] / Expected reference array, read only
    afActual   : ARRAY[1..64] OF REAL;   // 实际值数组，回读侧，只读不写 [工程单位] / Actual readback array, read only
END_VAR
VAR_INPUT
    nCount  : INT := 1;                  // 参与比对项数 [项]，域 1 到 64，越界钳位 / Item count, 1 to 64, clamped
    fAbsTol : REAL := 0.01;              // 统一绝对容差 [工程单位]，负值取绝对值 / Absolute tolerance, negative values folded to positive
END_VAR
VAR_OUTPUT
    nDiffCount   : INT;                  // 超差项数 [项] / Number of out of tolerance items
    nFirstDiffIdx : INT;                 // 首个超差项下标，0 表示无超差 [索引] / First out of tolerance index, zero when none
    fMaxDev      : REAL;                 // 最大绝对偏差值，只统计有限项 [工程单位] / Maximum absolute deviation over finite items
    nMaxDevIdx   : INT;                  // 最大偏差所在下标，0 表示未计算 [索引] / Index of the maximum deviation
    bEqual       : BOOL;                 // 全部项在容差内且无非有限值为真 / All items within tolerance and finite
    bNonFinite   : BOOL;                 // 出现过非数或非有限项为真 / NaN or infinity encountered
    uErrorId     : UDINT;                // 事件码，0 表示无事件 / Event code, zero means none
    bValid       : BOOL;                 // 项数与容差落在可服务域内为真，容差回退不否定结果 / Count and tolerance serviceable, a tolerance fallback does not void the result
END_VAR
VAR
    nCountUse : INT;                     // 生效项数，钳位后的值 [项] / Effective item count after clamping
    fTolUse   : REAL;                    // 生效容差，已取绝对值并钳到最小容差 [工程单位] / Effective tolerance after normalisation
    fDev      : REAL;                    // 单项绝对偏差 [工程单位] / Per item absolute deviation
    fA        : REAL;                    // 当前期望值快照 [工程单位] / Expected value snapshot
    fB        : REAL;                    // 当前实际值快照 [工程单位] / Actual value snapshot
    bFinA     : BOOL;                    // 期望值有限性判定结果 / Expected value finiteness
    bFinB     : BOOL;                    // 实际值有限性判定结果 / Actual value finiteness
    nGuard    : DINT;                    // 循环守卫计数，防遍历失控 [次] / Loop guard counter
    i         : INT;                     // 遍历索引，1 起 [索引] / Loop index, one based
END_VAR
VAR CONSTANT
    DL_ITEM_MAX   : INT := 64;          // 项数上限 [项] / Item count limit
    DL_GUARD_MAX  : DINT := 128;        // 循环守卫上限，两倍于项数上限故正常不触发 [次] / Loop guard limit, twice the item limit
    DL_I_MIN      : INT := 1;           // 数组首下标 [索引] / First array index
    DL_TOL_MIN    : REAL := 1.0E-9;     // 最小容差，容差为零时回退到此值 [工程单位] / Minimum tolerance used as the fallback
    DL_FINITE_MAX : REAL := 3.4E38;     // 有限性判定上限，超过即视为无穷大 [工程单位] / Finiteness ceiling, beyond this counts as infinity
END_VAR

(*------------------------------------------------------------------------------
 * 段 1｜输出预置：任何路径下输出确定
 *      Pre-set outputs so that every path is deterministic
 *-----------------------------------------------------------------------------*)
FC_DL_ArrayDiffSummary := FALSE;
nDiffCount             := 0;
nFirstDiffIdx          := 0;
fMaxDev                := 0.0;
nMaxDevIdx             := 0;
bEqual                 := FALSE;
bNonFinite             := FALSE;
uErrorId               := 16#0000_0000;
bValid                 := TRUE;

(*------------------------------------------------------------------------------
 * 段 2｜项数钳位（边界 B1）：先夹到 1 到 64 再进循环
 *      Clamp the item count into one to sixty four before the loop
 *-----------------------------------------------------------------------------*)
nCountUse := nCount;
IF nCountUse < DL_I_MIN THEN
    nCountUse := DL_I_MIN;
    bValid    := FALSE;
    uErrorId  := 16#0001_0134;   // 项数过小，已钳到下限
ELSIF nCountUse > DL_ITEM_MAX THEN
    nCountUse := DL_ITEM_MAX;
    bValid    := FALSE;
    uErrorId  := 16#0001_0134;   // 项数过大，已钳到上限
END_IF

(*------------------------------------------------------------------------------
 * 段 3｜容差归一（边界 B2）：先拦非数，再取绝对值，再钳最小容差
 *      Normalise the tolerance: reject NaN, fold sign, apply the lower bound
 *-----------------------------------------------------------------------------*)
IF fAbsTol <> fAbsTol THEN
    fTolUse := DL_TOL_MIN;
    IF uErrorId = 16#0000_0000 THEN
        uErrorId := 16#0001_0135;   // 容差为非数，回退到最小容差
    END_IF
ELSE
    fTolUse := ABS(fAbsTol);
    IF (fTolUse < DL_TOL_MIN) OR (fTolUse > DL_FINITE_MAX) THEN
        fTolUse := DL_TOL_MIN;
        IF uErrorId = 16#0000_0000 THEN
            uErrorId := 16#0001_0135;   // 容差过小或非有限，回退到最小容差
        END_IF
    END_IF
END_IF

(*------------------------------------------------------------------------------
 * 段 4｜单趟比对（边界 B3/B4/B5）：有限项走容差，非有限项直接计超差
 *      Single pass: finite items use the tolerance, non finite ones count as bad
 *-----------------------------------------------------------------------------*)
i      := DL_I_MIN;
nGuard := 0;
WHILE (i <= nCountUse) AND (nGuard < DL_GUARD_MAX) DO
    nGuard := nGuard + 1;

    fA    := afExpected[i];
    fB    := afActual[i];
    bFinA := NOT ((fA <> fA) OR (ABS(fA) > DL_FINITE_MAX));
    bFinB := NOT ((fB <> fB) OR (ABS(fB) > DL_FINITE_MAX));

    IF bFinA AND bFinB THEN
        fDev := ABS(fA - fB);
        IF fDev > DL_FINITE_MAX THEN
            (* 两个有限值相减仍可能溢出为无穷：按非有限处置，绝不参与最大偏差竞争 *)
            (* Two finite values can still overflow: treat it as non finite, no contest *)
            bNonFinite := TRUE;
            nDiffCount := nDiffCount + 1;
            IF nFirstDiffIdx = 0 THEN
                nFirstDiffIdx := i;
            END_IF
            fDev := 0.0;
        ELSE
            IF fDev > fTolUse THEN
                nDiffCount := nDiffCount + 1;
                IF nFirstDiffIdx = 0 THEN
                    nFirstDiffIdx := i;
                END_IF
            END_IF
            (* 最大偏差对所有有限项竞争，并列时取先出现者 *)
            (* The maximum is contested by every finite item, ties keep the earlier one *)
            IF fDev > fMaxDev THEN
                fMaxDev    := fDev;
                nMaxDevIdx := i;
            END_IF
        END_IF
    ELSE
        bNonFinite := TRUE;
        fDev       := 0.0;
        nDiffCount := nDiffCount + 1;
        IF nFirstDiffIdx = 0 THEN
            nFirstDiffIdx := i;
        END_IF
    END_IF

    i := i + 1;
END_WHILE

(*------------------------------------------------------------------------------
 * 段 5｜结论合成：无超差且无非有限值才算一致
 *      Verdict: equal only when no difference and every item is finite
 *-----------------------------------------------------------------------------*)
bEqual := (nDiffCount = 0) AND (NOT bNonFinite);

(*------------------------------------------------------------------------------
 * 段 6｜收口：返回一致性结论，合法性由 bValid 单独表达
 *      Close out: return the verdict, legality is expressed by bValid
 *-----------------------------------------------------------------------------*)
FC_DL_ArrayDiffSummary := bEqual;
END_FUNCTION

(* ---- FC_DL_ArrayFindValue.st ---- *)
(*
  ==================================================================
  组件名 Component  : FC_DL_ArrayFindValue
  分类   Category   : DL_MathData
  前缀   Naming     : FC_DL_ ｜ b/n/u/f/t/e/st 类型前缀制（R265）
  码位   Code ID    : 16#0001_0662（故障级）
  版本   Version    : 1.0.0
  复杂度 Complexity  : 低
  功能   Purpose    : LREAL 数组无序线性查找：返回目标值首 / 末命中下标与命中
                      计数三口径；未命中以 -1 哨兵表达，供值定位、重复检测、
                      抽检核对类调用方使用。
  开源溯源 Origin    : 西门子 LGF V5.3.0 Data Handling 组「数组搜索」子族
                      「无序线性查找 + 首 / 末 / 计数三口径」功能分类借鉴
                      （只借骨不抄肉）；实现 clean-room，零代码复制。
  许可证 License    : MIT
  参考   Reference  : IEC 61131-3:2013 §6.6.1 比较 / FOR 遍历语义
  平台   Platform   : 纯 IEC 61131-3（FOR / ABS / 比较），三平台通用
  依赖   Depends    : 无（零委托、零库件）
  分工声明 Split     : FC_DL_ArraySliceCopy（段拷贝）/ FC_DL_ArrayFindExtreme
                      （极值定位）与本件互引；本件为「值 → 下标」正向查找，
                      极值族为「无目标值」扫描，职责不同（R216）。
  归属 Ownership     : 本件无 TYPE 声明；全部引脚为 IEC 标准原生类型。
  ------------------------------------------------------------------
  边界 Boundary     :
                      一 nCount 越域（< 1 或 > 256）判故障早退（禁空遍历与
                         越界下标）；fValue 非有限判故障早退（禁 NaN 参与
                         容差比较）——两场景出口组合完全相同（三个计数均
                         哨兵值 + bValid = FALSE），合并一码（反证句见码表）；
                      二 样本非有限口径（声明）：afData 中的非有限样本
                         （NaN / ±Inf）**跳过**，不计命中也不报错（数组整体
                         仍可部分有效）；目标值 fValue 非有限则不在此口径内，
                         按边界一判故障；
                      三 命中判定用容差：ABS(样本 - 目标) < 1.0E-6，禁用
                         = / <> 判等（浮点判等红线）；
                      四 未命中哨兵：nFirst = -1 且 nLast = -1 且 nHits = 0，
                         bValid = TRUE（查找本身成功，无命中不是故障）；
                      五 纯函数：无记忆量、无定时器、无边沿实例，每调用重算；
                      六 无全局、无外部变量、无物理地址。
  错误码 Codes      :
    16#0001_0662【故障级】nCount 越域（< 1 或 > 256）或目标值 fValue 非有限
  码位反证 Note     :
    0662 合并「计数越域」与「目标值非有限」的理由：两场景出口组合完全相同
    （nFirst = -1、nLast = -1、nHits = 0、bValid = FALSE），三组以内输出无法
    唯一还原该场景，按 R90 不另立码；未命中（边界四）出口 bValid = TRUE，
    与 0662 可由 bValid 唯一区分，不并入。
  验收 Acceptance   :
    算法已证（脚本）：未跑 ｜ 编译器已证（三平台）：未跑
    V1 数组 [5, 7, 5, 9]、目标 5 → nFirst 0 / nLast 2 / nHits 2
    V2 目标 8 → 三哨兵 -1 / -1 / 0、bValid = TRUE（未命中不是故障）
    V3 含 NaN 样本 [NaN, 5]、目标 5 → NaN 跳过、nFirst 1 / nHits 1
    V4 nCount = 0 → 码 0662 + 早退（禁空遍历）
    V5 nCount = 257 → 同码早退；V6 目标 NaN → 同码早退
    V7 单样本命中 → nFirst = nLast = 0、nHits 1
  修订记录 Revision  :
    2026-11-21  v1.0.0  R64 首版（批 1 · 序号 2，LGF Data Handling 数组搜索子族）
  ==================================================================
*)
FUNCTION FC_DL_ArrayFindValue : BOOL
VAR_IN_OUT
    afData : ARRAY[0..255] OF LREAL; // 数据序列 [工程单位]，只读 / the data series, read only
END_VAR
VAR_INPUT
    nCount : DINT := 0;    // 有效样本数入参 [个]，合法域 1..256 / the sample count, legal one to two hundred fifty six
    fValue : LREAL := 0.0; // 查找目标值 [工程单位]，必须有限 / the target value, must be finite
END_VAR
VAR_OUTPUT
    nFirst : DINT;  // 首个命中下标 [下标]，未命中 = -1 哨兵 / the first hit index, minus one when no hit
    nLast  : DINT;  // 末个命中下标 [下标]，未命中 = -1 哨兵 / the last hit index, minus one when no hit
    nHits  : DINT;  // 命中计数 [个] / the hit count
    bValid : BOOL;  // 结果可用 [-]（未命中也是可用结果）/ the result usable, a no hit is still usable
    eErr   : UDINT; // 错误码，0 = 正常 / the error code, zero is ok
    bError : BOOL;  // 故障标志（故障级码同拍置位，R45 配对）/ the fault flag raised with a fault level code
END_VAR
VAR
    k : DINT := 0; // 遍历索引 [下标] / the traversal index
END_VAR  // R64 结构补齐：VAR 段缺失的 END_VAR（门禁机械修复）
VAR CONSTANT
    DL_AFP_NMAX : DINT := 256;       // 数组容量上界 [个]，与数组容量一致 / the capacity aligned with the array
    DL_AFP_ONE  : DINT := 1;         // 整型一常量 [个] / the integer one constant
    DL_AFP_NOHIT: DINT := -1;        // 未命中哨兵 [下标] / the no hit sentinel index
    DL_AFP_ZERO : DINT := 0;         // 整型零常量 [个] / the integer zero constant
    DL_AFP_EQEPS: LREAL := 1.0E-6;   // 命中容差 [工程单位]，禁用 = / <> 判等 / the hit tolerance, plain equality operators are forbidden
END_VAR

// 段 1｜返回值与全部出口预置哨兵值（R45 四段式第一段）/ segment 1, the preset of the return and all outlets
FC_DL_ArrayFindValue := FALSE; // 返回值预置假 / preset the return false
nFirst := DL_AFP_NOHIT; // 首命中下标预置哨兵 -1 [下标] / preset the first hit to the sentinel
nLast := DL_AFP_NOHIT; // 末命中下标预置哨兵 -1 [下标] / preset the last hit to the sentinel
nHits := DL_AFP_ZERO; // 命中计数预置零 [个] / preset the hit count zero
bValid := FALSE; // 可用标志预置假 / preset the validity false
eErr := 16#0000_0000; // 错误码预置正常 / preset the code to ok
bError := FALSE; // 故障标志预置假 / preset the fault flag false

// 段 2｜入参域闸（边界一，早退禁空遍历与 NaN 比较）/ segment 2, the input domain gate
IF (nCount < DL_AFP_ONE) OR (nCount > DL_AFP_NMAX)
OR (fValue <> fValue) OR ((fValue - fValue) <> (fValue - fValue)) THEN // 计数越域或目标值非有限 / the count is out of the domain or the target is not finite
    eErr := 16#0001_0662; // 故障级：入参越域或目标非有限（出口同形合并一码，R90）/ fault grade under the merged code
    bError := TRUE; // 同拍置故障标志（R45 配对）/ raise the fault flag on the same scan
    bValid := FALSE; // 结果不可用 / the result is not usable
    RETURN; // 早退 / early return
END_IF

// 段 3｜线性查找遍历（边界二：非有限样本跳过；边界三：容差判等）/ segment 3, the linear search traversal
FOR k := DL_AFP_ZERO TO nCount - DL_AFP_ONE DO // 有界遍历（上界已证 ≤ 256）/ the bounded traversal with a proven ceiling
    IF (afData[k] = afData[k]) AND ((afData[k] - afData[k]) = (afData[k] - afData[k])) THEN // 有限样本才参与（非有限跳过口径）/ only a finite sample participates
        IF ABS(afData[k] - fValue) < DL_AFP_EQEPS THEN // 容差命中（浮点禁判等）/ a hit inside the tolerance
            nHits := nHits + DL_AFP_ONE; // 命中计数推进 [个] / advance the hit count
            IF nFirst = DL_AFP_NOHIT THEN // 首个命中（哨兵未动过才写）/ the first hit only when the sentinel is intact
                nFirst := k; // 记首命中下标 [下标] / record the first hit index
            END_IF
            nLast := k; // 末命中下标随遍历自然收敛 [下标] / the last hit index converges along the traversal
        END_IF
    END_IF
END_FOR

// 段 4｜统一出口（未命中不是故障，边界四）/ segment 4, the unified outlet
bValid := TRUE; // 查找流程走完即可用（含未命中）/ the search completed, usable even with no hit
FC_DL_ArrayFindValue := TRUE; // 返回成功 / return success
END_FUNCTION

(* ---- FC_DL_ArraySliceCopy.st ---- *)
(*
  ==================================================================
  组件名 Component  : FC_DL_ArraySliceCopy
  分类   Category   : DL_MathData
  前缀   Naming     : FC_DL_ ｜ b/n/u/f/t/e/st 类型前缀制（R265）
  码位   Code ID    : 16#0001_0666（故障级）
  版本   Version    : 1.0.0
  复杂度 Complexity  : 低
  功能   Purpose    : 数值数组段拷贝：把源数组的 [iStart, iStart + nLen - 1]
                      段整段拷入目标数组首段起（目标从下标 0 起承接），LREAL
                      主类型；供缓冲搬运、窗段提取、队列重组类调用方使用。
  开源溯源 Origin    : 西门子 LGF V5.3.0 Data Handling 组「定长缓冲搬运（无
                      动态内存）」分类学口径借鉴（R12 结论沿用，只借骨不抄
                      肉）；实现 clean-room，零代码复制。
  许可证 License    : MIT
  参考   Reference  : IEC 61131-3:2013 §6.6.4 FOR 遍历与数组语义
  平台   Platform   : 纯 IEC 61131-3（FOR / 数组 / 比较），三平台通用
  依赖   Depends    : 无（零委托、零库件）
  分工声明 Split     : FC_DL_ArrayFindValue（值 → 下标查找）与本件互引；
                      本件只做段搬运不改序、不查值；数组裁剪压缩类需求由
                      调用方以本件 + 移位组合（R216）。
  归属 Ownership     : 本件无 TYPE 声明；全部引脚为 IEC 标准原生类型。
  ------------------------------------------------------------------
  边界 Boundary     :
                      一 入参域闸（逐项点名，R272）：nSrcCount < 1 或 > 256 /
                         iStart < 0 或 > nSrcCount - 1 / nLen < 1 或
                         nLen > nSrcCount - iStart（源溢出）或 nLen > 256
                         （目标容量溢出）→ 故障级 0666 + nCopied = 0 +
                         bValid = FALSE + 早退（禁任何写回，目标数组保持
                         原样）；四类越域出口组合完全相同，合并一码
                         （反证句见码表）；
                      二 重叠自检（中转缓冲两段式）：本件先把源段整段读入
                         局部中转缓冲，再整段写回目标——afSrc 与 afDst 为
                         同一数组且区间重叠的别名调用也不产生撕裂 / 串写
                         （快照语义，真实可达路径：调用方传同一数组做
                         前移压缩）；此为机制性防重叠，非永假防御；
                      三 拷贝序：中转缓冲承接后按下标 0 起顺序写回，循环
                         上界由段 1 域闸证明 ≤ 256，越界不可达；
                      四 纯函数：无记忆量、无定时器、无边沿实例，每调用重算；
                      五 无除法；无全局、无外部变量、无物理地址。
  错误码 Codes      :
    16#0001_0666【故障级】入参越域：nSrcCount / iStart / nLen 任一越出
                         合法域（源溢出或目标容量溢出，禁任何写回）
  码位反证 Note     :
    0666 合并四类越域（计数 / 起点 / 源溢出 / 容量溢出）的理由：四场景出口
    组合完全相同（nCopied = 0、bValid = FALSE、目标数组零写回），三组以内
    输出无法唯一还原该场景，按 R90 不另立码。
  验收 Acceptance   :
    算法已证（脚本）：未跑 ｜ 编译器已证（三平台）：未跑
    V1 源 [1,2,3,4,5]、iStart = 2、nLen = 3 → 目标 [3,4,5]、nCopied = 3
    V2 iStart = 0、nLen = nSrcCount → 全量拷贝
    V3 nLen = nSrcCount - iStart + 1（源溢出）→ 码 0666 + 早退、目标原样
    V4 iStart = nSrcCount（起点越界）→ 同码早退
    V5 nSrcCount = 0 / 257 → 同码早退
    V6 别名调用：afSrc = afDst 同数组、源段与目标首段重叠 → 中转缓冲两段式
       无撕裂（V1 结果断言不变）
  修订记录 Revision  :
    2026-11-21  v1.0.0  R64 首版（批 2 · 序号 5，LGF Data Handling 段拷贝补口）
  ==================================================================
*)
FUNCTION FC_DL_ArraySliceCopy : BOOL
VAR_IN_OUT
    afSrc : ARRAY[0..255] OF LREAL; // 源数组 [工程单位]，允许与目标同数组（别名调用走中转缓冲）/ the source array, may alias the target, the staging buffer covers it
    afDst : ARRAY[0..255] OF LREAL; // 目标数组 [工程单位]，从下标 0 起承接 / the target array, receives from the index zero
END_VAR
VAR_INPUT
    nSrcCount: DINT := 0; // 源有效长度 [个]，合法域 1..256 / the source effective length, legal one to two hundred fifty six
    iStart   : DINT := 0; // 源段起点 [下标]，合法域 0..nSrcCount - 1 / the source segment start index
    nLen     : DINT := 0; // 拷贝长度 [个]，合法域 1..min(nSrcCount - iStart, 256) / the copy length
END_VAR
VAR_OUTPUT
    nCopied: DINT;  // 实际拷贝数 [个]，失败 = 0 / the copied count, zero on failure
    bValid : BOOL;  // 结果可用 [-] / the result usable flag
    eErr   : UDINT; // 错误码，0 = 正常 / the error code, zero is ok
    bError : BOOL;  // 故障标志（故障级码同拍置位，R45 配对）/ the fault flag raised with a fault level code
END_VAR
VAR
    k         : DINT := 0;               // 遍历索引 [下标] / the traversal index
    afStaging : ARRAY[0..255] OF LREAL;  // 中转缓冲 [工程单位]，两段式防重叠撕裂 / the staging buffer for the overlap safe two stage copy
END_VAR  // R64 结构补齐：VAR 段缺失的 END_VAR（门禁机械修复）
VAR CONSTANT
    DL_ASC_NMAX : DINT := 256; // 数组容量上界 [个]，与数组容量一致 / the capacity aligned with the array
    DL_ASC_ONE  : DINT := 1;   // 整型一常量 [个] / the integer one constant
    DL_ASC_ZERO : DINT := 0;   // 整型零常量 [个] / the integer zero constant
END_VAR

// 段 1｜返回值与全部出口预置安全值（R45 四段式第一段）/ segment 1, the preset of the return and all outlets
FC_DL_ArraySliceCopy := FALSE; // 返回值预置假 / preset the return false
nCopied := DL_ASC_ZERO; // 拷贝数预置零 [个] / preset the copied count zero
bValid := FALSE; // 可用标志预置假 / preset the validity false
eErr := 16#0000_0000; // 错误码预置正常 / preset the code to ok
bError := FALSE; // 故障标志预置假 / preset the fault flag false
FOR k := DL_ASC_ZERO TO DL_ASC_NMAX - DL_ASC_ONE DO // 中转缓冲预清零（有界遍历全容量）/ preset the staging buffer zero over the full capacity
    afStaging[k] := 0.0; // 缓冲槽位显式清零 [工程单位] / clear the staging slot explicitly
END_FOR

// 段 2｜入参域闸（边界一：四类越域逐项点名，禁任何写回）/ segment 2, the input domain gate, no writeback on any violation
IF (nSrcCount < DL_ASC_ONE) OR (nSrcCount > DL_ASC_NMAX)
OR (iStart < DL_ASC_ZERO) OR (iStart > nSrcCount - DL_ASC_ONE)
OR (nLen < DL_ASC_ONE) OR (nLen > nSrcCount - iStart) OR (nLen > DL_ASC_NMAX) THEN // 计数 / 起点 / 长度任一越域 / the count or the start or the length is out of the domain
    eErr := 16#0001_0666; // 故障级：入参越域（四场景出口同形合并一码，R90）/ fault grade under the merged code
    bError := TRUE; // 同拍置故障标志（R45 配对）/ raise the fault flag on the same scan
    bValid := FALSE; // 结果不可用 / the result is not usable
    RETURN; // 早退，目标数组零写回 / early return, the target untouched
END_IF

// 段 3｜中转缓冲承接源段（边界二：两段式第一段，读侧快照）/ segment 3, the staging buffer takes the source segment
FOR k := DL_ASC_ZERO TO nLen - DL_ASC_ONE DO // 有界遍历（上界已证 ≤ 256 且 ≤ 源余量）/ the bounded traversal with a proven ceiling
    afStaging[k] := afSrc[iStart + k]; // 源段读入缓冲 [工程单位]（快照语义）/ read the source segment into the staging buffer
END_FOR

// 段 4｜缓冲写回目标（边界二：两段式第二段，写侧顺序落位）/ segment 4, the staging buffer lands on the target
FOR k := DL_ASC_ZERO TO nLen - DL_ASC_ONE DO // 有界遍历（上界同段 3 已证）/ the bounded traversal with the same proven ceiling
    afDst[k] := afStaging[k]; // 缓冲整段写回目标首段 [工程单位] / land the staging segment onto the target head
END_FOR

// 段 5｜统一出口 / segment 5, the unified outlet
nCopied := nLen; // 实拷贝数出口 [个] / the copied count outlet
bValid := TRUE; // 结果可用 / the result is usable
FC_DL_ArraySliceCopy := TRUE; // 返回成功 / return success
END_FUNCTION

(* ---- FC_DL_ArraySumLreal.st ---- *)
(*
    组件名称 : FC_DL_ArraySumLreal
    所属子库 : DL_MathData
    当前版本 : 1.0.0
    兼 容 性 : CODESYS V3.5+ / TwinCAT 3 / 汇川 InoProShop；仅依赖 Standard.library
    功能描述 : 静态数组一次性求和与均值，带非有限样本剔除与有效样本计数出口。
              取舍 ①：非有限样本剔除而不是让它们污染和 —— 一个 NaN 进和，整条链条全变 NaN，
              而均值 NaN 在 HMI 上显示为空白或 0，现场会当成「测量值为零」，这是最危险的静默错误；
              剔除 + nValidCount + 信息码，三点合起来让「有几个样本是坏的」变成可观测量。
              取舍 ②：均值独立判零分母 —— nValidCount = 0 时不算均值，直接判故障；
              绝不输出 0 冒充「均值为零」。
              取舍 ③：元素数超上限按上限钳位而非拒算 —— 静态表越界声明是配置问题，
              能算多少算多少并发信息码告警，比整表拒算更有用（配方系数、标定表都属这类）。
              取舍 ④：与 FB_DL_SignalStatistics 的边界 —— 那件是流式窗口（跨周期状态），
              本件是静态表一次性求值，纯函数、无内部状态、同入参同结果，可直接放进表达式或 CASE 分支里用。
    开源溯源 : 原创实现（T0-4 变体线，统计族「静态表求值」缺位）。无外部源码参考，码位与分级 100% 自有。；本件为 IEC 61131-3 标准语义的道莅防御性实现（原创实现，零外部源码复制）。
    本文件内含 : FUNCTION FC_DL_ArraySumLreal（单 POU，无配套类型）
    依 赖 : 无 DL_ 内部依赖；Standard.library: 无
    红线自检 : R1 ✓ 零全局变量与外部变量 ｜ R2 ✓ 零物理 IO 地址
              R3 ✓ 纯 IEC 61131-3 ｜ R4 ✓ 元素数闸 + 非有限剔除 + 均值判零分母 + 累加溢出复检
              R5 ✓ 全变量中英双语同行注释 ｜ R6 N/A 纯函数无顺序状态机，无 CASE 可写
              R7 N/A 无定时器、无沿检测实例 ｜ R8 ✓ 数组上限、有限域、容差全常量化
    错误码   : 16#0001_044C [信息级] 部分非有限样本已剔除，和与均值仅基于有效样本，bValid = TRUE
               16#0001_044D [信息级] 元素数超上限已按上限钳位，bValid = TRUE
               16#0001_0390 [故障级] 元素数为负，返回 0，bValid = FALSE
               16#0001_0391 [故障级] 无有效样本（全部非有限），和与均值均返回 0，bValid = FALSE
               16#0001_0392 [故障级] 累加溢出（中间量非有限），返回 0，bValid = FALSE
    码位总账 : 16#0001_044C 用 / 16#0001_044D 用 ｜ 16#0001_0390 用 / 16#0001_0391 用 / 16#0001_0392 用
    遗留假设 : ① 非有限判据用「自比较为假判 NaN + 幅值越界判 INF」，为 IEEE 754 语义推导，未在 InoProShop 实测。
              ② 均值的除法在 nValidCount > 0 时进行，除数为 INT_TO_LREAL(≥1)，除零结构性不可能。
    修订历史 :
        2026-11-16  v1.0.0  首版，R21 批次 3 入库
*)
FUNCTION FC_DL_ArraySumLreal : LREAL
VAR_INPUT
    nCount          : INT;    // 有效元素数，0~DL_ARRAY_MAX；超上限按上限钳位，负数判故障 [个] / number of valid elements, clamped above the bound and rejected below zero [count]
END_VAR
VAR_IN_OUT
    afData          : ARRAY[0..DL_ARRAY_MAX] OF LREAL;   // 定长数组，下标 ≥ nCount 的元素不参与 [工程单位] / fixed array, entries at or above nCount are ignored [engineering unit]
END_VAR
VAR_OUTPUT
    eErr            : UDINT;  // 错误码，0=正常；16#0001_04XX 信息级 / 16#0001_03XX 故障级 / error id, 0=ok
    bError          : BOOL;   // 故障级标志，eErr 落 16#0001_03XX 时为 TRUE / fault flag, TRUE on fault-level eErr
    bValid          : BOOL;   // 和与均值是否可用 / sum and mean usable flag
    fMean           : LREAL;  // 均值 = 和 / 有效样本数，无有效样本时为 0 [工程单位] / mean of the valid samples, zero when none is valid [engineering unit]
    nValidCount     : INT;    // 剔除非有限样本后的有效样本数 [个] / number of valid samples after the non-finite ones were dropped [count]
END_VAR
VAR
    nEff            : INT;    // 实际遍历元素数（钳位后）[个] / effective element count after clamping [count]
    nIdx            : INT;    // 数组游标 [个] / array cursor [count]
    nDropped        : INT;    // 被剔除的非有限样本数 [个] / number of dropped non-finite samples [count]
    fSum            : LREAL;  // 累加和 [工程单位] / running sum [engineering unit]
    fSample         : LREAL;  // 当前样本值 [工程单位] / current sample [engineering unit]
    bSampleFin      : BOOL;   // 当前样本是否有限 / whether the current sample is finite
END_VAR
VAR CONSTANT
    DL_ARRAY_MAX        : INT := 255;                          // 数组下标上限 [个] / array upper index [count]
    DL_ARRAY_NONE       : INT := 0;                            // 零元素哨兵，均值判零分母用 [个] / zero element sentinel guarding the mean division [count]
    DL_LREAL_MAX_FINITE : LREAL := 1.7976931348623157E308;     // LREAL 最大有限值 [无量纲] / largest finite LREAL [dimensionless]
    DL_LREAL_ZERO       : LREAL := 0.0;                        // 零哨兵 [工程单位] / zero sentinel [engineering unit]
    DL_ERR_NONE         : UDINT := 16#0000_0000;               // 无故障 / no error
END_VAR

// 段 1｜返回值与错误状态预置 / segment 1, preset the return value and the error state
FC_DL_ArraySumLreal := DL_LREAL_ZERO;   // 故障缺省返回 0 / fault default returns zero
eErr         := DL_ERR_NONE;            // 预置无错误 / preset no error
bError       := FALSE;                  // 预置无故障 / preset no fault
bValid       := FALSE;                  // 预置结果不可用 / preset unusable
fMean        := DL_LREAL_ZERO;          // 预置均值 0 / preset the mean to zero
nValidCount  := 0;                      // 预置有效样本 0 / preset the valid count to zero
nDropped     := 0;                      // 预置剔除数 0 / preset the dropped count to zero
fSum         := DL_LREAL_ZERO;          // 累加器清零 / clear the accumulator
nEff         := nCount;                 // 先按请求数占位 / start from the requested count

// 段 2｜元素数闸：负值判故障，超上限钳位并告警 / segment 2, count gate, reject negatives and clamp above the bound
IF nCount < DL_ARRAY_NONE THEN
    eErr   := 16#0001_0390;             // 元素数为负（故障级）/ negative element count, fault level
    bError := TRUE;                     // 置故障标志 / raise the fault flag
    RETURN;                             // 返回 0，bValid 保持 FALSE / return zero, bValid stays FALSE
END_IF
IF nCount > DL_ARRAY_MAX THEN
    nEff := DL_ARRAY_MAX;               // 钳到上限，能算多少算多少 / clamp to the bound and evaluate what is available
    eErr := 16#0001_044D;               // 元素数超上限已钳位（信息级，不置 bError）/ count clamped, info level
END_IF

// 段 3｜单遍求和：非有限样本剔除并计数，不污染和 / segment 3, single pass sum with non-finite samples dropped
IF nEff > DL_ARRAY_NONE THEN
    FOR nIdx := 0 TO nEff - 1 DO
        fSample    := afData[nIdx];                                                     // 取当前样本 / fetch the sample
        bSampleFin := (fSample = fSample) AND (ABS(fSample) <= DL_LREAL_MAX_FINITE);     // 自比较判 NaN，幅值判 INF / self compare for NaN, magnitude for INF
        IF bSampleFin THEN
            fSum := fSum + fSample;     // 只累加有效样本 / accumulate only valid samples
        ELSE
            nDropped := nDropped + 1;   // 剔除并计数 / drop and count
        END_IF
    END_FOR
END_IF
nValidCount := nEff - nDropped;         // 有效样本数 = 遍历数 − 剔除数 / valid count equals the visited minus the dropped

// 段 4｜剔除提示（先置者保留：超上限码若已占则不覆盖）/ segment 4, drop hint, never overwriting an existing code
IF (nDropped > 0) AND (eErr = DL_ERR_NONE) THEN
    eErr := 16#0001_044C;               // 非有限样本已剔除（信息级）/ non-finite samples dropped, info level
END_IF

// 段 5｜累加溢出复检：中间量非有限即溢出 / segment 5, overflow re-check on the accumulator
IF (fSum <> fSum) OR (ABS(fSum) > DL_LREAL_MAX_FINITE) THEN
    FC_DL_ArraySumLreal := DL_LREAL_ZERO;   // 溢出不给伪值 / never emit a pseudo value on overflow
    eErr   := 16#0001_0392;                // 累加溢出（故障级）/ accumulation overflow, fault level
    bError := TRUE;                        // 置故障标志 / raise the fault flag
    RETURN;                                // bValid 保持 FALSE / bValid stays FALSE
END_IF

// 段 6｜无有效样本闸：均值绝不靠除零得出 / segment 6, no valid sample gate, the mean never comes out of a division by zero
IF nValidCount = DL_ARRAY_NONE THEN
    FC_DL_ArraySumLreal := DL_LREAL_ZERO;   // 和仍为 0 / the sum stays zero
    fMean  := DL_LREAL_ZERO;               // 均值不计算，置 0 / the mean is not computed
    eErr   := 16#0001_0391;                // 无有效样本（故障级）/ no valid sample, fault level
    bError := TRUE;                        // 置故障标志 / raise the fault flag
    RETURN;                                // bValid 保持 FALSE / bValid stays FALSE
END_IF

// 段 7｜出口 / segment 7, exit
FC_DL_ArraySumLreal := fSum;                               // 输出和 / publish the sum
fMean := fSum / INT_TO_LREAL(nValidCount);                 // 除数恒 ≥ 1，结构性安全 / the divisor is at least one by construction
bValid := TRUE;                                            // 结果可用 / the results are usable
END_FUNCTION

(* ---- FC_DL_AsciiFrameParse.st ---- *)
(*
  ==================================================================
  组件名 Component  : FC_DL_AsciiFrameParse
  分类   Category   : DL_MathData
  复杂度 Complexity  : 中
  版本   Version    : 1.0.0
  功能   Purpose    : ASCII 仪表帧解析。STX(16#02)/ETX(16#03) 定界 + 长度闸
                      + 可选校验。载荷校验模式：载荷末两字符为十六进制校验
                      和（前部载荷字符 hex 值之和模 256），bChkEn = TRUE 时
                      逐字符 hex 解码比对。OSCAT Network ASCII 帧族语义
                      clean-room，与 FC_DL_ModbusRtuFrameCheck 二进制帧分工。
  来源   Source     : T1-3-oscat-network（ASCII 帧族公开语义）
  溯源   Origin     : STX/ETX 定界与 LRC 校验为公开工业语义，clean-room 自研
                      实现，未复制 OSCAT 或任何厂商私有库源码。
  平台   Platform   : 纯 IEC 61131-3（Standard.library: LEN / MID / LEFT /
                      RIGHT / FIND，'$02' '$03' 为 IEC 标准 $ 转义）
  分工声明 Split     : 与 FC_DL_ModbusRtuFrameCheck 分工——后者做二进制 RTU
                      帧校验，本件做 ASCII 可打印帧解析。
  作者   Author     : 道莅代码库 · PLC 编程专家（R59）
  ------------------------------------------------------------------
  边界 Boundary     :
                      一 结构闸：长度 ∈ [5..255]（STX + 载荷 ≥1 + 校验 2 +
                         ETX）、首字符 = STX、末字符 = ETX、ETX 唯一（FIND
                         定位 = 末位），任一不满足置 bError；
                      二 校验闸（bChkEn）：载荷含非 hex 字符或和模 256 ≠ 校
                         和 → bBadChk（信息级），bValid 随之降假；
                      三 非有限无涉（纯整数与串操作，无除零/浮点风险）；
                      四 无全局变量、无外部变量声明、无物理地址寻址。
  修订记录 Revision  :
    2026-11-21  v1.0.0  R59 首版（批 2 · 序号 7）
  ==================================================================
*)

FUNCTION FC_DL_AsciiFrameParse : BOOL
VAR_INPUT
    sFrame : STRING(255) := ''; // 原始帧串（含 STX/ETX）[-] / the raw frame string with the delimiters
    bChkEn : BOOL := FALSE;     // 载荷校验使能（末两字符 hex 校验和）[-] / the payload checksum enable
END_VAR
VAR_OUTPUT
    sPayload : STRING(255) := ''; // 载荷输出（不含 STX/ETX/校验段，校验使能时）/ the payload outlet, without the delimiters and the checksum when enabled
    nPayLen  : DINT  := 0;  // 载荷长度 [字符] / the payload length
    bValid   : BOOL := FALSE; // 解析受理且校验通过（校验未使能时仅结构）[-] / the parsed and verified flag
    bBadChk  : BOOL := FALSE; // 校验不匹配或载荷非 hex（信息级，仅校验使能时判定）[-] / the checksum mismatch, informational
    bError   : BOOL := FALSE; // 结构故障标志（定界/长度闸）[-] / the structure fault flag
END_VAR
VAR CONSTANT
    DL_AFP_STX    : STRING(1) := '$02'; // 帧头 STX（IEC $ 转义）/ the STX delimiter
    DL_AFP_ETX    : STRING(1) := '$03'; // 帧尾 ETX（IEC $ 转义）/ the ETX delimiter
    DL_AFP_HEXTAB : STRING(16) := '0123456789ABCDEF'; // hex 字符表（FIND 解码）/ the hex table for the FIND decoding
    DL_AFP_LENMIN : DINT := 5;  // 最小帧长（STX+1+2+ETX）[字符] / the min frame length
    DL_AFP_LENMAX : DINT := 255; // 最大帧长（库串上限）[字符] / the max frame length
END_VAR
VAR
    nLen   : DINT; // 帧长 [字符] / the frame length
    nEtx   : DINT; // ETX 定位（FIND 结果）[位] / the ETX position by the FIND
    sCh    : STRING(1); // 单字符工作量 [-] / the one char work value
    nPos   : DINT;  // hex 表命中位（0 = 非法）[位] / the hex table hit, zero means illegal
    nSum   : DINT;  // 载荷 hex 值累加和 [无量纲] / the payload hex value sum
    nChk   : DINT;  // 末两字符校验和值 [无量纲] / the trailing checksum value
    nI     : DINT;  // 载荷遍历索引 [字符] / the payload loop index
    nDataLen: DINT; // 数据段长度（载荷减校验两字符）[字符] / the data length, the payload minus two
    sHead  : STRING(1); // 首字符工作量 [-] / the first char work value
    sTail  : STRING(1); // 末字符工作量 [-] / the last char work value
    sChk   : STRING(2); // 校验段工作量 [-] / the checksum slice work value
END_VAR

// 段 1｜返回值与输出预置（四段式第一段，R45）/ segment 1, preset the return and the outputs
FC_DL_AsciiFrameParse := FALSE; // 受理预置假 / preset the accepted false
sPayload := ''; // 载荷预置空 / preset the payload empty
nPayLen := 0; // 载荷长预置零 / preset the payload length zero
bValid := FALSE; // 有效预置假 / preset the valid false
bBadChk := FALSE; // 校验不匹配预置假 / preset the checksum flag false
bError := FALSE; // 故障预置假 / preset the fault false

// 段 2｜结构闸（定界 + 长度 + ETX 唯一性，边界一）/ segment 2, the structure gates
nLen := LEN(sFrame); // 取帧长 / take the frame length
IF (nLen < DL_AFP_LENMIN) OR (nLen > DL_AFP_LENMAX) THEN // 长度闸 / the length gate
    bError := TRUE; // 置故障 / raise the fault
    RETURN; // 早退 / return early
END_IF
sHead := LEFT(sFrame, 1); // 取首字符 / take the first char
sTail := RIGHT(sFrame, 1); // 取末字符 / take the last char
IF (sHead <> DL_AFP_STX) OR (sTail <> DL_AFP_ETX) THEN // 定界闸 / the delimiter gate
    bError := TRUE; // 置故障 / raise the fault
    RETURN; // 早退 / return early
END_IF
nEtx := FIND(sFrame, DL_AFP_ETX); // ETX 定位 / locate the ETX
IF nEtx <> nLen THEN // ETX 非末位（帧内混入 ETX）/ the ETX not at the tail
    bError := TRUE; // 置故障 / raise the fault
    RETURN; // 早退 / return early
END_IF

// 段 3｜载荷提取与校验判定（校验使能时载荷末两字符为 hex 校验和，边界二）/ segment 3, the payload extraction and the checksum
IF bChkEn THEN // 校验使能模式 / the checksum enabled mode
    nDataLen := nLen - 5; // 数据段长 = 帧长 - STX - ETX - 校验 2 字符 / the data length
    sPayload := MID(sFrame, nDataLen, 2); // 取数据段（跳过 STX 与校验两字符）/ take the data slice
    sChk := MID(sFrame, 2, nDataLen + 1); // 取校验两字符 / take the two checksum chars
    nSum := 0; // 和清零 / clear the sum
    FOR nI := 1 TO nDataLen DO // 逐数据字符 hex 累加 / per data char hex sum
        sCh := MID(sPayload, 1, nI); // 取单字符 / take one char
        nPos := FIND(DL_AFP_HEXTAB, sCh); // hex 表命中 / the hex table hit
        IF nPos = 0 THEN // 非 hex 字符 / a non hex char
            bBadChk := TRUE; // 置校验不匹配（信息级）/ raise the mismatch, informational
        ELSE // 合法 hex / a legal hex
            nSum := nSum + (nPos - 1); // 累加 hex 值 / accumulate the value
        END_IF
    END_FOR
    nPos := FIND(DL_AFP_HEXTAB, MID(sChk, 1, 1)); // 校验高位解码 / decode the high nibble
    IF nPos = 0 THEN // 非法 / illegal
        bBadChk := TRUE; // 置不匹配 / raise the mismatch
    ELSE // 合法 / legal
        nChk := (nPos - 1) * 16; // 高位 ×16 / the high times sixteen
        nPos := FIND(DL_AFP_HEXTAB, MID(sChk, 1, 2)); // 校验低位解码 / decode the low nibble
        IF nPos = 0 THEN // 非法 / illegal
            bBadChk := TRUE; // 置不匹配 / raise the mismatch
        ELSE // 合法 / legal
            nChk := nChk + (nPos - 1); // 低位并入 / add the low
            IF (nSum MOD 256) <> nChk THEN // 和模 256 比对 / the modulo compare
                bBadChk := TRUE; // 校验不匹配 / the mismatch
            END_IF
        END_IF
    END_IF
    nPayLen := nDataLen; // 载荷长出口（数据段口径）/ the payload length outlet
ELSE // 校验未使能：整段载荷直通 / the checksum disabled, the whole payload
    sPayload := MID(sFrame, nLen - 2, 2); // 取 STX 与 ETX 之间 / take between the delimiters
    nPayLen := nLen - 2; // 载荷长出口 / the payload length outlet
    IF nPayLen < 1 THEN // 零载荷防御（长度闸已保下限 5，纵深）/ the empty payload defense in depth
        bError := TRUE; // 置故障 / raise the fault
        RETURN; // 早退 / return early
    END_IF
END_IF

// 段 4｜统一出口（校验使能时 bValid = 结构通过 AND 校验通过）/ segment 4, the unified outlet
bValid := (NOT bError) AND (NOT bBadChk); // 受理判据 / the accept verdict
FC_DL_AsciiFrameParse := bValid; // 受理标志 / the accepted flag
END_FUNCTION

(* ---- FC_DL_AsinDegChk.st ---- *)
(*==============================================================================
 * 名称 : FC_DL_AsinDegChk —— 反正弦 → 角度（输入钳位 [-1,1]，越界仍按钳位计算）
 * 分类 / 前缀 / 版本 : DL_MathData / FC_DL_ / 1.0.0
 * 溯源 : 开源语义参考（OSCAT/AixOCAT 族，MIT）或 clean-room IEC 实现，未复制源码
 * 平台 : 纯 IEC 61131-3
 * 功能说明 : 返回 asin(x) 的角度制结果 [-90,90]。输入越出 [-1,1] 时钳位到
 *            边界后仍按钳位值计算（bValid=FALSE、eErr 置码提示越界），不产生
 *            NaN。恒等式 asin(x)=atan2(x, sqrt(1-x^2))（弧度）转角度输出，
 *            纯 ATAN2/SQRT 内联实现，无库内跨件依赖。
 *            边界处理：输入非有限（NaN/±Inf）置 eErr 返回 0.0（不钳位计算）。
 * 错误码 : 16#0001_1B0C = 输入越出 [-1,1]（已钳位计算），或输入非有限（NaN/±Inf）
 *          eErr=0 且 bValid=TRUE 表示输入在域内、返回值可用
 * 状态机 : R6 标注 N/A（纯函数无顺序状态，以本节替代 ELSE 兜底）
 * 红线 : R1/R2/R3 ✓ 零全局/零IO/纯IEC ｜ R4 ✓ 非有限拦截/域钳位防 NaN ｜ R10 ✓ 标准转换 ｜ R11 ✓ 分号收尾 ｜ R15 ✓ 无保留字撞名
 * 修订记录 : 2026-11-23 v1.0.0 首次入库（R76）
 *============================================================================*)
FUNCTION FC_DL_AsinDegChk : LREAL
VAR_INPUT
    fX : LREAL;    // 正弦值输入 [-1,1]，越界钳位 / sine value input, clamped into [-1,1]
END_VAR
VAR_OUTPUT
    eErr   : UDINT;    // 故障码，0=正常，1B0C=越界钳位或非有限 / error code
    bError : BOOL;     // TRUE=本件发生故障 / TRUE when fault occurred
    bValid : BOOL;     // TRUE=输入在域内且返回值可用 / TRUE when input in domain and result usable
END_VAR
VAR
    _x   : LREAL;      // 钳位后的输入 [无量纲] / clamped input
    _fR  : LREAL;      // 弧度制反正弦结果 [rad] / arcsine result in radians
END_VAR

FC_DL_AsinDegChk := 0.0;                     // 返回值预设 0.0 / preset return to zero
eErr   := 16#0000_0000;                      // 故障码清零 / clear error code
bError := FALSE;                             // 故障标志清零 / clear error flag
bValid := TRUE;                              // 预设输出可用 / preset valid flag

IF (fX <> fX) OR ((fX - fX) <> (fX - fX)) THEN    // NaN 或 ±Inf / NaN or infinite
    eErr   := 16#0001_1B0C;                  // 置非有限故障码 / set non-finite code
    bError := TRUE;                          // 置故障标志 / set error flag
    bValid := FALSE;                         // 返回值不可用 / return not usable
    RETURN;                                  // 返回 0.0 / return zero
END_IF

_x := fX;                                    // 取输入 / take input
IF _x > 1.0 THEN                             // 上越界钳位 / clamp upper
    _x := 1.0;                               // 钳到 +1 / clamp to +1
    eErr   := 16#0001_1B0C;                  // 置越界码 / set out-of-domain code
    bError := TRUE;                          // 置故障标志 / set error flag
    bValid := FALSE;                         // 提示越界（仍按钳位值出结果）/ flag clamped compute
ELSIF _x < -1.0 THEN                         // 下越界钳位 / clamp lower
    _x := -1.0;                              // 钳到 -1 / clamp to -1
    eErr   := 16#0001_1B0C;                  // 置越界码 / set out-of-domain code
    bError := TRUE;                          // 置故障标志 / set error flag
    bValid := FALSE;                         // 提示越界（仍按钳位值出结果）/ flag clamped compute
END_IF

_fR := ATAN2(_x, SQRT(1.0 - _x * _x));       // asin(x)=atan2(x,sqrt(1-x^2))，弧度 / arcsine via atan2
FC_DL_AsinDegChk := _fR * 180.0 / 3.14159265358979323846;    // 弧度转角度 / radians to degrees

END_FUNCTION

(* ---- FC_DL_AsinEx.st ---- *)
(*
    FC_DL_AsinEx —— 反正弦防御包装（定义域 [-1,1] 域闸钳位 + NaN 拦截）
    ------------------------------------------------------------------
    分类      : DL_MathData / Math-Trig
    前缀      : FC_DL_
    版本      : 1.0.0
    溯源      : IEC 61131-3 标准语义的道莅防御性实现
                （内部委托平台内建函数，外围统一错误码/钳位/双语文档；
                  未复制任何闭源厂商源码，参考实现仅限 MIT/Apache 许可）
    平台      : 纯 IEC 61131-3，CODESYS / TwinCAT / InoProShop 通用
    作者      : 道莅代码库 · PLC编程专家（R15）
    ------------------------------------------------------------------
    功能说明  : 求输入的反正弦，返回值域 [-pi/2, pi/2]。定义域闸门先行：
                NaN 输入拦截返回 0.0 并置 16#0001_016D；定义域 [-1,1] 之外（含
                无穷）钳位到 ±1 并置 16#0001_016D，bValid=FALSE 但仍返回钳位后的
                计算结果（±pi/2）供降级使用；域内委托内建 ASIN，边界值
                ±1 为合法输入直接通过；结果再做 NaN 复检兜底。
    错误码    : 0000 正常 / 16#0001_016D 入参越界（NaN 已归零，或域外已钳位到 ±1）
    修订记录  : 2026-11-16 v1.0.0 首次入库（R15）
*)
FUNCTION FC_DL_AsinEx : LREAL
VAR_INPUT
    lrIn : LREAL; // 输入实数 [无量纲]，定义域 [-1,1] / input real value [dimensionless], domain minus 1 to plus 1
END_VAR
VAR_OUTPUT
    eErr : UDINT; // 错误码，0=正常，1=入参越界（已钳位/归零） / error id, 0=ok, 1=input out of domain, clamped or zeroed
    bError   : BOOL; // 是否出错，eErr 非 0 时为 TRUE / error flag, TRUE when eErr is nonzero
    bValid   : BOOL; // 输出是否有效可用，钳位/归零降级时为 FALSE / output valid, FALSE for clamped or zeroed degraded results
END_VAR
VAR
    lrUse : LREAL; // 钳位后的实际计算入参 [无量纲] / clamped value actually fed to the kernel [dimensionless]
END_VAR
VAR CONSTANT
    DL_AS_DOM : LREAL := 1.0; // 定义域边界 [无量纲]，闭区间 / domain bound [dimensionless], closed interval
END_VAR

// 段 1｜返回值与错误状态预置，任何早退路径不留脏码 / segment 1, preset return value and error states
FC_DL_AsinEx := 0.0; // 返回值预置安全值 0.0 / preset return to safe value 0.0
eErr    := 16#0000_0000; // 错误码预置正常 / preset error id to ok
bError      := FALSE; // 错误标志预置无错 / preset error flag to FALSE
bValid      := TRUE; // 有效标志预置可用 / preset valid flag to TRUE

// 段 2｜NaN 拦截：自不等判据，归零早退，不进内核 / segment 2, NaN interception by self-inequality, zeroed early exit
IF lrIn <> lrIn THEN
    eErr := 16#0001_016D; // 信息级：输入 NaN，已归零 / informational, NaN input, zeroed
    bError   := TRUE; // 置错误标志 / raise error flag
    bValid   := FALSE; // 输出不可用 / output invalid
    RETURN; // 返回预置安全值 0.0 / return preset safe value 0.0
END_IF

// 段 3｜定义域闸门：域外（含无穷）钳位到 ±1，仍返回钳位后结果 / segment 3, domain gate, out-of-domain including infinity clamped to plus or minus 1 with result still returned
IF lrIn > DL_AS_DOM THEN
    lrUse    := DL_AS_DOM; // 上越界钳位 +1 / upper overflow clamped to plus 1
    eErr := 16#0001_016D; // 信息级：域外已钳位 / informational, out of domain clamped
    bError   := TRUE; // 置错误标志 / raise error flag
    bValid   := FALSE; // 钳位结果非真实值 / clamped result is not the true value
ELSIF lrIn < -DL_AS_DOM THEN
    lrUse    := -DL_AS_DOM; // 下越界钳位 -1 / lower overflow clamped to minus 1
    eErr := 16#0001_016D; // 信息级：域外已钳位 / informational, out of domain clamped
    bError   := TRUE; // 置错误标志 / raise error flag
    bValid   := FALSE; // 钳位结果非真实值 / clamped result is not the true value
ELSE
    lrUse := lrIn; // 域内直通（±1 边界合法） / in-domain pass-through, boundary plus or minus 1 legal
END_IF

// 段 4｜委托内建 ASIN / segment 4, delegation to built-in ASIN
FC_DL_AsinEx := ASIN(lrUse); // 委托内建 ASIN 内核 / delegate to built-in ASIN kernel

// 段 5｜结果 NaN 复检兜底（防御纵深，正常路径不可达） / segment 5, result NaN recheck as defense in depth
IF FC_DL_AsinEx <> FC_DL_AsinEx THEN
    FC_DL_AsinEx := 0.0; // 兜底安全值 / bottom-line safe value
    IF eErr = 16#0000_0000 THEN
        eErr := 16#0001_016D; // 首事件优先置码 / first-event priority code
        bError   := TRUE; // 置错误标志 / raise error flag
        bValid   := FALSE; // 输出不可用 / output invalid
    END_IF
END_IF
END_FUNCTION

(* ---- FC_DL_AsinSafe.st ---- *)
(*
    FC_DL_AsinSafe —— 反正弦 Safe 族防御包装（域钳位 + bClamped 显式标志 + 委托内建）
    ------------------------------------------------------------------
    分类      : DL_MathData / Math-Trig
    前缀      : FC_DL_
    版本      : 1.0.0
    来源标签  : iec-std-wrapper（T0）
    溯源      : IEC 61131-3 标准语义的道莅防御性实现
                （内部委托平台内建 ASIN，外围钳位/错误码/双语文档；
                  未复制任何闭源厂商源码）
    平台      : 纯 IEC 61131-3，CODESYS / TwinCAT / InoProShop 通用
    分工声明  : 与存量 FC_DL_AsinEx 分工——AsinEx 为码位族（16#0001_016D 口径），
                本件为 Safe 族样板（bClamped 显式钳位标志 + 16#0002 子带码位），
                两件并存服务不同调用方约定，算法内核同为内建 ASIN 委托。
    作者      : 道莅代码库 · PLC 编程专家（R57）
    ------------------------------------------------------------------
    功能说明  : 求输入的反正弦，返回值域 [-pi/2, pi/2]。四段式防御（R45）：
                NaN 双判据拦截归零早退；|x|>1（含无穷）钳到 ±1 并置 bClamped
                仍返回钳位结果供降级；域内委托内建 ASIN；结果 NaN 复检兜底。
    错误码    : 0000 正常 / 16#0002_0001 入参非有限已归零 / 16#0002_0002 域外已钳位
    修订记录  : 2026-11-21 v1.0.0 首次入库（R57 批 2 · 序号 6）
*)
FUNCTION FC_DL_AsinSafe : LREAL
VAR_INPUT
    lrIn : LREAL; // 输入实数 [无量纲]，定义域 [-1,1] / input real value [dimensionless], domain minus one to plus one
END_VAR
VAR_OUTPUT
    eErr     : UDINT; // 错误码，0 = 正常 / error code, zero is ok
    bError   : BOOL;  // 出错标志，eErr 非 0 时为真 / error flag, true when eErr is nonzero
    bValid   : BOOL;  // 结果是否为真实值，钳位/归零降级时为假 / the result is the true value, false when degraded
    bClamped : BOOL;  // 本次调用发生定义域钳位 [-] / a domain clamp happened this call
END_VAR
VAR
    lrUse : LREAL; // 钳位后的实际计算入参 [无量纲] / the clamped value fed to the kernel [dimensionless]
END_VAR
VAR CONSTANT
    DL_ASN_DOM : LREAL := 1.0; // 定义域边界 [无量纲]，闭区间 / the domain bound [dimensionless], closed interval
END_VAR

// 段 1｜返回值与错误状态预置安全值（四段式第一段，R45）/ segment 1, preset the return and error states
FC_DL_AsinSafe := 0.0; // 返回值预置安全值 0.0 / preset the return to the safe zero
eErr     := 16#0000_0000; // 错误码预置正常 / preset the code to ok
bError   := FALSE; // 错误标志预置假 / preset the error flag false
bValid   := TRUE; // 有效标志预置真 / preset the valid flag true
bClamped := FALSE; // 钳位标志预置假 / preset the clamp flag false

// 段 2｜非有限拦截（双判据）：命中不调内建直接早退 / segment 2, the non finite interception, early exit without the kernel
IF (lrIn <> lrIn) OR ((lrIn - lrIn) <> (lrIn - lrIn)) THEN // NaN 或无穷 / NaN or infinity
    eErr   := 16#0002_0001; // 信息级：输入非有限已归零 / informational, a non finite input zeroed
    bError := TRUE; // 置错误标志 / raise the error flag
    bValid := FALSE; // 输出不可用 / the output void
    RETURN; // 返回预置安全值 0.0 / return the preset safe zero
END_IF

// 段 3｜定义域闸门：域外钳到 ±1 并置 bClamped，仍返回钳位结果 / segment 3, the domain gate, clamped to plus or minus one with the flag raised
IF lrIn > DL_ASN_DOM THEN // 上越界（含正无穷，已被段 2 拦截故此处为有限值）/ above the bound
    lrUse    := DL_ASN_DOM; // 钳到 +1 / clamp to plus one
    eErr     := 16#0002_0002; // 信息级：域外已钳位 / informational, clamped
    bError   := TRUE; // 置错误标志 / raise the error flag
    bValid   := FALSE; // 钳位结果非真实值 / the clamped result is not the true value
    bClamped := TRUE; // 置钳位标志 / raise the clamp flag
ELSIF lrIn < -DL_ASN_DOM THEN // 下越界 / below the bound
    lrUse    := -DL_ASN_DOM; // 钳到 -1 / clamp to minus one
    eErr     := 16#0002_0002; // 信息级：域外已钳位 / informational, clamped
    bError   := TRUE; // 置错误标志 / raise the error flag
    bValid   := FALSE; // 钳位结果非真实值 / the clamped result is not the true value
    bClamped := TRUE; // 置钳位标志 / raise the clamp flag
ELSE // 域内直通（±1 边界合法）/ inside the domain, the boundary legal
    lrUse := lrIn; // 直通 / passthrough
END_IF

// 段 4｜委托内建 ASIN（禁重实现数学内核）/ segment 4, delegation to the built-in ASIN
FC_DL_AsinSafe := ASIN(lrUse); // 委托内建内核 / delegate to the built-in kernel

// 段 5｜结果 NaN 复检兜底（防御纵深，正常路径不可达）/ segment 5, the result recheck as defense in depth
IF (FC_DL_AsinSafe <> FC_DL_AsinSafe) OR ((FC_DL_AsinSafe - FC_DL_AsinSafe) <> (FC_DL_AsinSafe - FC_DL_AsinSafe)) THEN // 结果非有限 / a non finite result
    FC_DL_AsinSafe := 0.0; // 兜底安全值 / the bottom-line safe value
    IF eErr = 16#0000_0000 THEN // 首事件优先置码 / the first event keeps the code
        eErr   := 16#0002_0001; // 信息级：结果非有限已归零 / informational, a non finite result zeroed
        bError := TRUE; // 置错误标志 / raise the error flag
        bValid := FALSE; // 输出不可用 / the output void
    END_IF
END_IF
END_FUNCTION

(* ---- FC_DL_Atan2Deg.st ---- *)
(*==============================================================================
 * 名称 : FC_DL_Atan2Deg —— 四象限反正切 → 角度 [0,360)（原点双重合防护）
 * 分类 / 前缀 / 版本 : DL_MathData / FC_DL_ / 1.0.0
 * 溯源 : 开源语义参考（OSCAT/AixOCAT 族，MIT）或 clean-room IEC 实现，未复制源码
 * 平台 : 纯 IEC 61131-3
 * 功能说明 : 返回 atan2(fY, fX) 的角度制结果并归一到 [0,360)（数学域
 *            (-180,180] 中负角加 360°）。两输入同时为 0 时方向无定义，
 *            返回 0.0、bValid=FALSE 并置 eErr。
 *            边界处理：任一输入非有限（NaN/±Inf）置 eErr 返回 0.0；fX=0 且
 *            fY≠0 的 ±90° 轴向情形由 ATAN2 数值语义原生支持，无需特判。
 * 错误码 : 16#0001_1B0E = fX 与 fY 同时为 0（方向无定义），或输入非有限（NaN/±Inf）
 *          eErr=0 且 bValid=TRUE 表示返回值可用
 * 状态机 : R6 标注 N/A（纯函数无顺序状态，以本节替代 ELSE 兜底）
 * 红线 : R1/R2/R3 ✓ 零全局/零IO/纯IEC ｜ R4 ✓ 非有限拦截/原点零向量防护 ｜ R10 ✓ 标准转换 ｜ R11 ✓ 分号收尾 ｜ R15 ✓ 无保留字撞名
 * 修订记录 : 2026-11-23 v1.0.0 首次入库（R76）
 *============================================================================*)
FUNCTION FC_DL_Atan2Deg : LREAL
VAR_INPUT
    fY : LREAL;    // 纵向分量 [工程单位] / vertical component
    fX : LREAL;    // 横向分量 [工程单位] / horizontal component
END_VAR
VAR_OUTPUT
    eErr   : UDINT;    // 故障码，0=正常，1B0E=零向量或非有限 / error code
    bError : BOOL;     // TRUE=本件发生故障 / TRUE when fault occurred
    bValid : BOOL;     // TRUE=返回值可用 / TRUE when return value is usable
END_VAR
VAR
    _d : LREAL;        // 角度中间值 [度] / angle intermediate in degrees
END_VAR

FC_DL_Atan2Deg := 0.0;                       // 返回值预设 0.0 / preset return to zero
eErr   := 16#0000_0000;                      // 故障码清零 / clear error code
bError := FALSE;                             // 故障标志清零 / clear error flag
bValid := TRUE;                              // 预设输出可用 / preset valid flag

IF (fY <> fY) OR ((fY - fY) <> (fY - fY))    // fY 非有限 / fY is NaN or infinite
   OR (fX <> fX) OR ((fX - fX) <> (fX - fX)) THEN    // fX 非有限 / fX is NaN or infinite
    eErr   := 16#0001_1B0E;                  // 置非有限故障码 / set non-finite code
    bError := TRUE;                          // 置故障标志 / set error flag
    bValid := FALSE;                         // 返回值不可用 / return not usable
    RETURN;                                  // 返回 0.0 / return zero
END_IF

IF (fY = 0.0) AND (fX = 0.0) THEN            // 零向量：方向无定义 / zero vector: no direction
    eErr   := 16#0001_1B0E;                  // 置零向量故障码 / set zero-vector code
    bError := TRUE;                          // 置故障标志 / set error flag
    bValid := FALSE;                         // 返回值不可用 / return not usable
    FC_DL_Atan2Deg := 0.0;                   // 返回 0.0（契约约定）/ return zero per contract
    RETURN;                                  // 提前收口 / early exit
END_IF

_d := ATAN2(fY, fX) * 180.0 / 3.14159265358979323846;    // 四象限反正弦转角度 / atan2 to degrees
IF _d < 0.0 THEN                             // 负角修正到 [0,360) / fold negative into [0,360)
    _d := _d + 360.0;                        // 加一整圈 / add one turn
END_IF

FC_DL_Atan2Deg := _d;                        // 回写 [0,360) 方向角 / write back direction

END_FUNCTION

(* ---- FC_DL_Atan2Ex.st ---- *)
(*
    FC_DL_Atan2Ex —— 四象限反正切防御包装（y,x 双入参 + 双零定义 + NaN/Inf 复检）
    ------------------------------------------------------------------
    分类      : DL_MathData / Math-Trig
    前缀      : FC_DL_
    版本      : 1.0.0
    溯源      : IEC 61131-3 标准语义的道莅防御性实现
                （内部委托平台内建函数，外围统一错误码/钳位/双语文档；
                  未复制任何闭源厂商源码，参考实现仅限 MIT/Apache 许可）
    平台      : 纯 IEC 61131-3，CODESYS / TwinCAT / InoProShop 通用
    作者      : 道莅代码库 · PLC编程专家（R15）
    ------------------------------------------------------------------
    功能说明  : 求四象限反正切 ATAN2(y,x)，返回 (-pi, pi]。处理次序写死：
                ① NaN 拦截归零早退；② 双零判据（|x|<1.0E-12 且 |y|<1.0E-12）
                返回 0.0 置 16#0001_017E 信息码（bError=TRUE、bValid=FALSE，需上层
                注意）；③ 近零 x 轴判向返回 ±pi/2；④ x>0 委托 ATAN(y/x)；
                ⑤ x<0 按 y 符号加/减 pi；⑥ IF 链尾无条件 ELSE 兜底返回
                0.0 置 16#0001_024B；⑦ 结果 NaN 复检兜底（拦截 Inf/Inf 组合毒值）。
                除法分支均在 |x|>=1.0E-12 保证下执行，无除零风险。
    错误码    : 0000 正常 / 16#0001_017C 入参越界 / 16#0001_017E 双零输入无定义（信息级） / 16#0001_024B 结果不可表示（兜底）
    修订记录  : 2026-11-16 v1.0.0 首次入库（R15）
*)
FUNCTION FC_DL_Atan2Ex : LREAL
VAR_INPUT
    lrY : LREAL; // 纵分量 [无量纲]，任意有限值或 NaN/无穷 / y component [dimensionless], any finite value or NaN/inf
    lrX : LREAL; // 横分量 [无量纲]，任意有限值或 NaN/无穷 / x component [dimensionless], any finite value or NaN/inf
END_VAR
VAR_OUTPUT
    eErr : UDINT; // 错误码，0=正常，4=双零输入，5=结果不可表示 / error id, 0=ok, 4=double zero input, 5=result not representable
    bError   : BOOL; // 是否出错，eErr 非 0 时为 TRUE / error flag, TRUE when eErr is nonzero
    bValid   : BOOL; // 输出是否有效可用，降级/兜底时为 FALSE / output valid, FALSE for degraded or fallback results
END_VAR
VAR
    lrOut : LREAL; // 计算结果中间量 [rad] / intermediate result [rad]
END_VAR
VAR CONSTANT
    DL_A2_EPS     : LREAL := 1.0E-12; // 双零/近零判据 [无量纲] / double-zero and near-zero threshold [dimensionless]
    DL_A2_PI      : LREAL := 3.1415926535897932; // 圆周率 [rad] / pi [rad]
    DL_A2_PI2     : LREAL := 1.5707963267948966; // 圆周率一半 [rad] / half pi [rad]
    DL_A2_MAXREAL : LREAL := 1.7976931348623157E308; // 双精度有限极值 [无量纲] / double precision finite max [dimensionless]
END_VAR

// 段 1｜返回值与错误状态预置，任何早退路径不留脏码 / segment 1, preset return value and error states
lrOut      := 0.0; // 结果中间量预置安全值 / preset intermediate result to safe value
eErr   := 16#0000_0000; // 错误码预置正常 / preset error id to ok
bError     := FALSE; // 错误标志预置无错 / preset error flag to FALSE
bValid     := TRUE; // 有效标志预置可用 / preset valid flag to TRUE

// 段 2｜NaN 拦截：任一分量为 NaN 一律归零早退 / segment 2, NaN interception, either component NaN zeroed early exit
IF (lrY <> lrY) OR (lrX <> lrX) THEN
    eErr := 16#0001_017C; // 信息级：输入 NaN，已归零 / informational, NaN input, zeroed
    bError   := TRUE; // 置错误标志 / raise error flag
    bValid   := FALSE; // 输出不可用 / output invalid
    FC_DL_Atan2Ex := lrOut;
    RETURN;
END_IF

// 段 3｜四象限 IF/ELSIF 判定链，链尾含无条件 ELSE 兜底 / segment 3, quadrant if-elsif chain with unconditional else fallback
IF (ABS(lrX) < DL_A2_EPS) AND (ABS(lrY) < DL_A2_EPS) THEN
    lrOut    := 0.0; // 双零输入按约定返回 0.0 / double-zero input returns 0.0 by convention
    eErr := 16#0001_017E; // 信息级：双零输入无定义 / informational, double-zero input undefined
    bError   := TRUE; // 置错误标志以示上层注意 / raise error flag for upper layer attention
    bValid   := FALSE; // 约定值非真实角度 / conventional value is not a true angle
ELSIF ABS(lrX) < DL_A2_EPS THEN
    IF lrY > 0.0 THEN
        lrOut := DL_A2_PI2; // 正 y 轴 +pi/2 / positive y axis plus half pi
    ELSIF lrY < 0.0 THEN
        lrOut := -DL_A2_PI2; // 负 y 轴 -pi/2 / negative y axis minus half pi
    ELSE
        lrOut    := 0.0; // 理论不可达兜底 / theoretically unreachable fallback
        eErr := 16#0001_024B; // 结果不可表示 / result not representable
        bError   := TRUE; // 置错误标志 / raise error flag
        bValid   := FALSE; // 输出不可用 / output invalid
    END_IF
ELSIF lrX > 0.0 THEN
    lrOut := ATAN(lrY / lrX); // 右半平面一/四象限 / right half plane quadrants 1 and 4, division guarded by the epsilon branch
ELSIF lrX < 0.0 THEN
    IF lrY >= 0.0 THEN
        lrOut := ATAN(lrY / lrX) + DL_A2_PI; // 左上半平面二象限 / upper-left half plane quadrant 2
    ELSE
        lrOut := ATAN(lrY / lrX) - DL_A2_PI; // 左下半平面三象限 / lower-left half plane quadrant 3
    END_IF
ELSE
    lrOut    := 0.0; // 无条件兜底分支，理论不可达 / unconditional fallback branch, theoretically unreachable
    eErr := 16#0001_024B; // 结果不可表示 / result not representable
    bError   := TRUE; // 置错误标志 / raise error flag
    bValid   := FALSE; // 输出不可用 / output invalid
END_IF

// 段 4｜结果 NaN 复检兜底：拦截 Inf/Inf 等组合产生的毒值 / segment 4, result NaN recheck, intercepts poisoned values from combinations like Inf over Inf
IF lrOut <> lrOut THEN
    lrOut := 0.0; // 兜底安全值 / bottom-line safe value
    IF eErr = 16#0000_0000 THEN
        eErr := 16#0001_024B; // 结果不可表示 / result not representable
        bError   := TRUE; // 置错误标志 / raise error flag
        bValid   := FALSE; // 输出不可用 / output invalid
    END_IF
END_IF

// 段 5｜有限性钳位复检与输出 / segment 5, finiteness clamp recheck and output
IF lrOut > DL_A2_MAXREAL THEN
    lrOut := DL_A2_MAXREAL; // 超极值钳位（防御纵深） / clamp beyond-extreme value, defense in depth
ELSIF lrOut < -DL_A2_MAXREAL THEN
    lrOut := -DL_A2_MAXREAL; // 超负极值钳位（防御纵深） / clamp beyond-negative-extreme value, defense in depth
END_IF
FC_DL_Atan2Ex := lrOut; // 输出四象限角 [rad] / output the quadrant angle
END_FUNCTION

(* ---- FC_DL_AtanEx.st ---- *)
(*
    FC_DL_AtanEx —— 反正切防御包装（全实数域 + NaN/无穷拦截降级）
    ------------------------------------------------------------------
    分类      : DL_MathData / Math-Trig
    前缀      : FC_DL_
    版本      : 1.0.0
    溯源      : IEC 61131-3 标准语义的道莅防御性实现
                （内部委托平台内建函数，外围统一错误码/钳位/双语文档；
                  未复制任何闭源厂商源码，参考实现仅限 MIT/Apache 许可）
    平台      : 纯 IEC 61131-3，CODESYS / TwinCAT / InoProShop 通用
    作者      : 道莅代码库 · PLC编程专家（R15）
    ------------------------------------------------------------------
    功能说明  : 求输入的反正切，全实数域合法，返回值域 (-pi/2, pi/2)。
                NaN 输入拦截返回 0.0 并置 16#0001_0177；正无穷按极限口径返回
                pi/2、负无穷返回 -pi/2，均置 16#0001_0177 且 bValid=FALSE 降级；
                有限域内直接委托内建 ATAN；结果再做 NaN 复检兜底，全程
                不输出 NaN/Inf。
    错误码    : 0000 正常 / 16#0001_0177 入参越界（NaN 已归零，或无穷已取极限值降级）
    修订记录  : 2026-11-16 v1.0.0 首次入库（R15）
*)
FUNCTION FC_DL_AtanEx : LREAL
VAR_INPUT
    lrIn : LREAL; // 输入实数 [无量纲]，全实数域 / input real value [dimensionless], full real domain
END_VAR
VAR_OUTPUT
    eErr : UDINT; // 错误码，0=正常，1=入参越界（NaN/无穷降级） / error id, 0=ok, 1=input out of domain (NaN or infinity degraded)
    bError   : BOOL; // 是否出错，eErr 非 0 时为 TRUE / error flag, TRUE when eErr is nonzero
    bValid   : BOOL; // 输出是否有效可用，降级时为 FALSE / output valid, FALSE for degraded results
END_VAR
VAR CONSTANT
    DL_AT_MAXREAL : LREAL := 1.7976931348623157E308; // 双精度有限极值 [无量纲]，超界判无穷 / double precision finite max [dimensionless], beyond treated as infinity
    DL_AT_PI2     : LREAL := 1.5707963267948966; // 圆周率一半 [rad]，无穷极限值 / half pi [rad], limit value at infinity
END_VAR

// 段 1｜返回值与错误状态预置，任何早退路径不留脏码 / segment 1, preset return value and error states
FC_DL_AtanEx := 0.0; // 返回值预置安全值 0.0 / preset return to safe value 0.0
eErr    := 16#0000_0000; // 错误码预置正常 / preset error id to ok
bError      := FALSE; // 错误标志预置无错 / preset error flag to FALSE
bValid      := TRUE; // 有效标志预置可用 / preset valid flag to TRUE

// 段 2｜NaN 拦截：自不等判据，归零早退，不进内核 / segment 2, NaN interception by self-inequality, zeroed early exit
IF lrIn <> lrIn THEN
    eErr := 16#0001_0177; // 信息级：输入 NaN，已归零 / informational, NaN input, zeroed
    bError   := TRUE; // 置错误标志 / raise error flag
    bValid   := FALSE; // 输出不可用 / output invalid
    RETURN; // 返回预置安全值 0.0 / return preset safe value 0.0
END_IF

// 段 3｜无穷降级闸：按极限口径返回 ±pi/2 并置 16#0001_0177 / segment 3, infinity degradation gate, limit value plus or minus half pi returned with code 1
IF lrIn > DL_AT_MAXREAL THEN
    FC_DL_AtanEx := DL_AT_PI2; // 正无穷极限 +pi/2 / plus infinity limit plus half pi
    eErr     := 16#0001_0177; // 信息级：输入无穷，已取极限值 / informational, infinite input, limit value returned
    bError       := TRUE; // 置错误标志 / raise error flag
    bValid       := FALSE; // 降级输出 / degraded output
    RETURN;
ELSIF lrIn < -DL_AT_MAXREAL THEN
    FC_DL_AtanEx := -DL_AT_PI2; // 负无穷极限 -pi/2 / minus infinity limit minus half pi
    eErr     := 16#0001_0177; // 信息级：输入无穷，已取极限值 / informational, infinite input, limit value returned
    bError       := TRUE; // 置错误标志 / raise error flag
    bValid       := FALSE; // 降级输出 / degraded output
    RETURN;
END_IF

// 段 4｜有限域内委托内建 ATAN / segment 4, finite domain delegation to built-in ATAN
FC_DL_AtanEx := ATAN(lrIn); // 委托内建 ATAN 内核 / delegate to built-in ATAN kernel

// 段 5｜结果 NaN 复检兜底（防御纵深，正常路径不可达） / segment 5, result NaN recheck as defense in depth
IF FC_DL_AtanEx <> FC_DL_AtanEx THEN
    FC_DL_AtanEx := 0.0; // 兜底安全值 / bottom-line safe value
    IF eErr = 16#0000_0000 THEN
        eErr := 16#0001_0177; // 首事件优先置码 / first-event priority code
        bError   := TRUE; // 置错误标志 / raise error flag
        bValid   := FALSE; // 输出不可用 / output invalid
    END_IF
END_IF
END_FUNCTION
